(* IEC 61131-3 sources: daoli-st-library/DL_Process (part 51) *)

(* ---- FB_DL_ShiftHandoverCheck.st ---- *)
(*
  ==================================================================
  组件名 Component  : FB_DL_ShiftHandoverCheck
  分类   Category   : DL_Process
  复杂度 Complexity  : 中
  版本   Version    : 1.0.1
  功能   Purpose    : 班次交接检查。交接开始沿取运行快照（产量与报警计数），
                      交接窗 tHandover 内逐条确认未决事项，全部确认即置完成单拍
                      bHandoverDone；窗到期仍有未决项则升级故障码并转未完成态。
  来源   Source     : self-std（IEC 61131-3 标准时序 + 交接业务语义自研）
  溯源   Origin     : 班次交接检查为公开生产管理语义，道莅 clean-room 自研实现，
                      未复制任何厂商私有库源码。
  平台   Platform   : 纯 IEC 61131-3（TON / R_TRIG / 比较），三平台通用
  分工声明 Split     : 与 FB_DL_ShiftMonthReport（报表属主）与 FB_DL_ChangeoverSequence
                      （产品换型属主）双向互补——本件只做交接时点的检查与确认闭环，
                      不出报表、不做换型顺控、不改动生产计数本体。
  作者   Author     : 道莅代码库 · PLC 编程专家（R60）
  归属 Ownership     : E_DL_HandoverPhase 属主为本文件（全库唯一定义，R264）；
                      引用件只引用不重声明（D13 返修补行）。
  接口偏离声明       : nProdCnt / nAlarmCnt 为 UDINT 却沿用 n 前缀（D10 返修登记
                      例外，R200）：沿用派单既有引脚名不改，避免破坏调用方接口；
                      族内新件一律用 u 前缀。
  ------------------------------------------------------------------
  边界 Boundary     :
                      一 零长窗显式分支（R253）：tHandover ≤ 0 判组态非法故障码，
                         不进交接相（禁靠比较算子隐式分流）；
                      二 同拍竞态让位于合法事件（R275）：交汇段先消化本拍确认沿，
                         再消化窗口到期迁移——到期拍恰有确认沿时按确认处理，
                         不在同拍升级超窗码；
                      三 进入/退出条件逐条取反对偶（R259）：进入 = 开始沿 + 使能 +
                         窗合法 + 无锁存；退出 = 全确认（完成）/ 窗口到期（升级）/
                         失能（弃用）/ 复位沿（清锁存）四条并列；
                      四 快照「最近一次」类出口纳入复位清单（R243）：nSnapProd 与
                         nSnapAlarm 在复位沿一并清零；
                      五 单拍输出 bHandoverDone 统一出口段每拍先预置 FALSE、
                         分支只写 TRUE（R256）；
                      六 使能 bEnable = FALSE 时语义为「弃用本轮交接」（转空闲，
                         不锁存、不出单拍）——R191 声明行；
                      七 故障解除路径：eFault 相由复位沿迁回空闲并清锁存与快照
                         （bReset 为输入引脚，恒可达，R152 自证）。
  错误码   Codes    :
    16#0005_0620【信息级】交接窗内尚有未决事项（逐拍重算，不锁存）
    16#0005_0621【故障级】交接窗时长非法（≤0），组态非法，锁存至复位沿
    16#0005_0622【故障级】交接窗到期仍未全部确认，升级未完成故障，锁存至复位沿
  验收   Acceptance :
    算法已证（脚本）：未跑 ｜ 编译器已证（三平台）：未跑
    V1 3 项未决、窗内 3 个确认沿 → bHandoverDone 单拍、无故障
    V2 窗到期仅确认 2/3 → 码 0622、eFault、未完成
    V3 tHandover = T#0S → 首拍即码 0621，不进交接相
  修订记录 Revision  :
    2026-11-21  v1.0.0  R60 首版（批 3 · 序号 12）
    2026-11-21  v1.0.1  R61 返修：D7 增 _nPendingLock，仅 eIdle 迁入沿赋值，
                        判据与注释对齐（R259）；D10 n 前缀 UDINT 字段登记
                        例外；D13 补 E_DL_HandoverPhase 属主行
  ==================================================================
*)

TYPE E_DL_HandoverPhase :
(
    eIdle  := 0,  // 空闲：等交接开始沿 / idle, waiting for the start edge
    eWait  := 10, // 等待：交接窗内逐条确认 / waiting for the item confirmations inside the window
    eFault := 20  // 故障：窗非法或到期未完成，锁存待复位 / fault, an illegal window or an unfinished overrun, latched
);
END_TYPE

FUNCTION_BLOCK FB_DL_ShiftHandoverCheck
VAR_INPUT
    bEnable      : BOOL := TRUE;       // 使能，FALSE 时弃用本轮交接（边界六）/ the enable, false discards the round
    bStart       : BOOL := FALSE;      // 交接开始电平，上升沿取快照 / the start level, the rising edge takes the snapshot
    bConfirmItem : BOOL := FALSE;      // 未决事项确认电平，上升沿确认一条 / the item confirmation level, each rising edge confirms one item
    bReset       : BOOL := FALSE;      // 复位沿：清锁存与快照并回空闲 / the reset edge, clears the latch and the snapshot
    tHandover    : TIME := T#10M;      // 交接窗时长 [毫秒]，必须 > 0 / the handover window, must be positive
    nPendingItems : DINT := 3;         // 未决事项条数 [条]，合法域 0..64 / the pending item count, legal from zero to sixty four
    nProdCnt     : UDINT := 0;         // 当前班次产量计数 [件] / the production count of the shift
    nAlarmCnt    : UDINT := 0;         // 当前班次报警计数 [次] / the alarm count of the shift
END_VAR
VAR_OUTPUT
    bRunning       : BOOL := FALSE;               // 交接窗口进行中 [-] / the handover in progress flag
    bHandoverDone  : BOOL := FALSE;               // 交接完成单拍脉冲 [-] / the handover done one shot pulse
    nConfirmedCnt  : DINT := 0;                   // 已确认条数 [条] / the confirmed item count
    nSnapProd      : UDINT := 0;                  // 交接开始时刻的产量快照 [件] / the production snapshot at the start edge
    nSnapAlarm     : UDINT := 0;                  // 交接开始时刻的报警快照 [次] / the alarm snapshot at the start edge
    eState         : E_DL_HandoverPhase;          // 主状态机当前态 [状态] / the current state of the main machine
    bError         : BOOL := FALSE;               // 故障锁存位 [-] / the latched fault bit
    eErr           : UDINT := 16#0000_0000;       // 错误码，0 = 正常 / the error code, zero is ok
END_VAR
VAR
    _bInit      : BOOL := FALSE;                                 // 首拍初始化标志（R310）/ the first scan flag
    _eState     : E_DL_HandoverPhase := E_DL_HandoverPhase.eIdle; // 内部状态寄存器，段 4 唯一写点 / the internal state register, single writer
    _bDone      : BOOL := FALSE;                                 // 完成单拍内部位，段 1 预清段 6 映射 / the internal done bit, preset then mapped
    _nConfirmed : DINT := 0;                                     // 已确认条数副本 / the confirmed count copy
    _nPending   : DINT := 0;                                     // 未决条数钳位工作副本（逐拍重算，仅供迁入沿快照，D7 返修）/ the clamped pending work copy, recomputed every scan
    _nPendingLock : DINT := 0;                                   // 本轮未决条数锁定值（仅 eIdle 迁入沿赋值，D7 返修，R259）/ the locked pending count, assigned only on the idle entry edge
    _uSnapProd  : UDINT := 0;                                    // 产量快照副本 / the production snapshot copy
    _uSnapAlarm : UDINT := 0;                                    // 报警快照副本 / the alarm snapshot copy
    _bFault     : BOOL := FALSE;                                 // 故障锁存副本（仅复位沿清除）/ the fault latch copy
    _bCfgBad    : BOOL := FALSE;                                 // 组态非法标记（逐拍重算）[-] / the configuration fault flag
    _bIncomplete : BOOL := FALSE;                                // 未确认标记（逐拍重算）[-] / the unconfirmed flag
    rtStart     : R_TRIG;                                        // 开始沿实例，段 0 无条件刷新 / the start edge instance
    rtConfirm   : R_TRIG;                                        // 确认沿实例，段 0 无条件刷新 / the confirmation edge instance
    rtReset     : R_TRIG;                                        // 复位沿实例，段 0 无条件刷新 / the reset edge instance
    tonWindow   : TON;                                           // 交接窗定时器，段 0 无条件刷新 / the handover window timer
END_VAR
VAR CONSTANT
    DL_SHC_ITMAX : DINT := 64; // 未决事项上界 [条] / the pending item bound
END_VAR

// 段 0｜沿检测与交接窗定时器无条件周期刷新（禁入分支，R7；IN 串故障锁存门控，FB50-1）/ segment 0, the unconditional refresh with the latch gate
rtStart(CLK := bStart); // 开始沿 / the start edge
rtConfirm(CLK := bConfirmItem); // 确认沿 / the confirmation edge
rtReset(CLK := bReset); // 复位沿 / the reset edge
tonWindow(IN := (_eState = E_DL_HandoverPhase.eWait) AND (NOT _bFault), PT := tHandover); // 交接窗：仅等待相且无锁存时计时 / the window timing only in the waiting phase

// 段 1｜首拍初始化与单拍标志预清（仅单拍标志入清单，R32 FB32-1；R256）/ segment 1, the first scan init and the one shot preset
IF NOT _bInit THEN // 首拍一拍 / the first scan
    _bInit := TRUE; // 置首拍标志 / raise the first scan flag
    _nConfirmed := 0; // 已确认条数显式清零 / clear the confirmed count explicitly
    _nPending := 0; // 未决条数显式清零 / clear the pending count explicitly
    _nPendingLock := 0; // 未决锁定值显式清零（D7 返修）/ clear the locked pending count explicitly
    _uSnapProd := 0; // 产量快照显式清零 / clear the production snapshot explicitly
    _uSnapAlarm := 0; // 报警快照显式清零 / clear the alarm snapshot explicitly
    _bFault := FALSE; // 故障锁存显式清零 / clear the fault latch explicitly
    _eState := E_DL_HandoverPhase.eIdle; // 状态显式落空闲 / place the state to idle explicitly
END_IF
_bDone := FALSE; // 完成单拍预清零 / preset the done pulse false
_bCfgBad := FALSE; // 组态非法标记预清零 / preset the configuration flag false
_bIncomplete := FALSE; // 未确认标记预清零 / preset the unconfirmed flag false

// 段 2｜组态域闸（零长窗显式分支，边界一；未决条数越域钳位）/ segment 2, the configuration gate with the explicit zero length branch
IF tHandover <= T#0S THEN // 零长窗：非法组态 / a zero length window, an illegal configuration
    _bCfgBad := TRUE; // 置组态非法标记 / raise the configuration flag
    _bFault := TRUE; // 锁存故障（段 5 迁移相）/ latch the fault, the segment five migrates the phase
END_IF
IF nPendingItems < 0 THEN // 条目数为负（域下界硬限）/ a negative item count
    _nPending := 0; // 按零条处理（无未决即完成）/ treat as zero, an immediate completion
ELSIF nPendingItems > DL_SHC_ITMAX THEN // 条目数越上界 / above the bound
    _nPending := DL_SHC_ITMAX; // 钳到上界 / clamp to the bound
ELSE // 域内 / inside the domain
    _nPending := nPendingItems; // 原值接管 / take the value as is
END_IF

// 段 3｜本拍确认沿预消化（R275：合法事件先于窗口到期迁移消化，段序在段 4 之前）/ segment 3, the confirmation edge pre digest ahead of the window expiry
IF rtConfirm.Q AND (_eState = E_DL_HandoverPhase.eWait) AND (NOT _bFault) THEN // 等待相内的确认沿 / a confirmation edge inside the waiting phase
    IF _nConfirmed < _nPendingLock THEN // 尚有未确认条目（判据用锁定值，D7 返修）/ items remain unconfirmed against the locked count
        _nConfirmed := _nConfirmed + 1; // 确认一条 / confirm one item
    ELSE // 已全部确认（多按的确认沿忽略）/ everything is confirmed, extra presses ignored
        _nConfirmed := _nPendingLock; // 计数饱和于锁定条目数 / saturate the count at the locked item count
    END_IF
END_IF

// 段 4｜主状态机（ENUM + CASE，ELSE 拦非法态；进入/退出逐条取反对偶，边界三）/ segment 4, the main machine with the paired entry and exit conditions
CASE _eState OF
    E_DL_HandoverPhase.eIdle: // 空闲相：等开始沿（条件：开始沿 + 使能 + 窗合法 + 无锁存）/ the idle phase
        IF rtStart.Q AND bEnable AND (tHandover > T#0S) AND (NOT _bFault) THEN // 迁入判据带全量闸位复检（R274）/ the entry with the full gate recheck
            _nConfirmed := 0; // 新一轮确认计数归零 / reset the confirmed count
            _uSnapProd := nProdCnt; // 取产量快照（最近一次类出口）/ take the production snapshot
            _uSnapAlarm := nAlarmCnt; // 取报警快照 / take the alarm snapshot
            _nPendingLock := _nPending; // 未决条数锁定（仅此迁入沿赋值，窗内改参不影响本轮判据，D7 返修）/ lock the pending count on this entry edge only
            _eState := E_DL_HandoverPhase.eWait; // 迁入等待相 / enter the waiting phase
        END_IF
    E_DL_HandoverPhase.eWait: // 等待相：四条退出（全确认 / 到期 / 失能 / 锁存）/ the waiting phase with four exits
        IF _nConfirmed >= _nPendingLock THEN // 退出条件一：全部确认（判据用锁定值，D7 返修）/ the first exit, everything confirmed against the locked count
            _bDone := TRUE; // 置完成单拍 / raise the done pulse
            _eState := E_DL_HandoverPhase.eIdle; // 迁回空闲 / back to idle
        ELSIF tonWindow.Q THEN // 退出条件二：窗口到期仍未全部确认（边界二：本拍确认沿已在段 3 消化）/ the second exit, the window expired unconfirmed
            _bIncomplete := TRUE; // 置未确认标记 / raise the unconfirmed flag
            _bFault := TRUE; // 锁存超窗故障（0622）/ latch the overrun fault
        ELSIF (NOT bEnable) OR _bFault THEN // 退出条件三：失能弃用或已锁存（前置条件消失）/ the third exit with the prerequisite gone
            _eState := E_DL_HandoverPhase.eIdle; // 迁回空闲（不锁存、不出单拍）/ back to idle without a latch or a pulse
        END_IF
    E_DL_HandoverPhase.eFault: // 故障相：锁存保持，等复位沿（解除可达，边界七）/ the fault phase held until the reset edge
        IF rtReset.Q THEN // 复位沿（复位作用域：清锁存 + 清快照 + 清累计量 + 迁相位）/ the reset with the declared scope
            _bFault := FALSE; // 清故障锁存 / clear the fault latch
            _nConfirmed := 0; // 清确认计数 / clear the confirmed count
            _nPendingLock := 0; // 清未决锁定值（复位作用域含锁定值，D7 返修）/ clear the locked pending count within the reset scope
            _uSnapProd := 0; // 清产量快照（R243 最近一次类出口入复位清单）/ clear the production snapshot
            _uSnapAlarm := 0; // 清报警快照 / clear the alarm snapshot
            _eState := E_DL_HandoverPhase.eIdle; // 故障相迁出边回空闲 / the exit edge back to idle
        END_IF
    ELSE // 非法枚举值拦截 / the illegal enumeration guard
        _eState := E_DL_HandoverPhase.eIdle; // 落回空闲 / force back to idle
        _bFault := TRUE; // 置故障锁存 / latch the fault
END_CASE

// 段 5｜故障锁存迁移闸（置于解除段之后防同拍抢迁，R258）/ segment 5, the fault latch to phase gate placed after the release
IF _bFault AND (_eState <> E_DL_HandoverPhase.eFault) THEN // 已锁存但不在故障相 / latched but not in the fault phase
    _eState := E_DL_HandoverPhase.eFault; // 迁入故障相 / enter the fault phase
END_IF

// 段 6｜统一出口（内部副本单点映射，R180；故障码锁存回放，R187）/ segment 6, the unified outlet
_bIncomplete := (_eState = E_DL_HandoverPhase.eWait) AND (_nConfirmed < _nPendingLock); // 未确认提示逐拍重算（判据用锁定值，D7 返修）/ the unconfirmed hint recomputed every scan against the locked count
bRunning := (_eState = E_DL_HandoverPhase.eWait); // 进行中出口 / the in progress outlet
bHandoverDone := _bDone; // 完成单拍出口 / the done pulse outlet
nConfirmedCnt := _nConfirmed; // 确认条数出口 / the confirmed count outlet
nSnapProd := _uSnapProd; // 产量快照出口 / the production snapshot outlet
nSnapAlarm := _uSnapAlarm; // 报警快照出口 / the alarm snapshot outlet
eState := _eState; // 状态出口 / the state outlet
bError := _bFault; // 故障位出口（与锁存同源）/ the fault bit outlet from the same latch
IF _bFault THEN // 故障锁存回放优先 / the latched fault replays first
    IF _bCfgBad THEN // 组态成因（独立码值，R190）/ the configuration cause with its own code
        eErr := 16#0005_0621; // 故障级：交接窗时长非法 / fault grade, the window length is illegal
    ELSE // 超窗成因 / the overrun cause
        eErr := 16#0005_0622; // 故障级：到期仍未全部确认 / fault grade, still unconfirmed at the expiry
    END_IF
ELSIF _bIncomplete THEN // 未确认提示（信息级，逐拍重算）/ the informational unconfirmed hint
    eErr := 16#0005_0620; // 信息级：尚有未决事项 / informational, items still pending
    bError := FALSE; // 信息级不置 bError（仅故障级置位，R45 配对口径）/ the informational code never raises the fault bit
ELSE // 无事件 / no event
    eErr := 16#0000_0000; // 正常 / ok
END_IF
END_FUNCTION_BLOCK

(* ---- FB_DL_ShiftMonthReport.st ---- *)
(*
  ==================================================================
  组件名 Component  : FB_DL_ShiftMonthReport
  分类   Category   : DL_Process
  版本   Version    : 1.0.0
  功能   Purpose    : 班次 / 月度窗口产量报表闸。班次结束脉冲到达时结算本班产量
                      （好品 / 废品 / 良率）并累加进月度窗口，同时打开报表闸
                      （等上位确认或超时自动关闸），关闸拍出报表完成脉冲。
                      月变更沿清月度累计与班次计数，实现「班次窗 + 月度窗」双窗一致。
  溯源   Origin     : 班次 / 月度报表闸为通用产量统计语义；本件为 clean-room 实现，
                      仅借鉴来源分类与参数域组织（来源标签 roadmap-p2-shift），
                      道莅原创设计，未复制任何闭源代码行。
  平台   Platform   : 纯 IEC 61131-3（R_TRIG / TON / UDINT / REAL，无私有库）
  作者   Author     : 道莅代码库 · PLC 编程专家（R55）
  ------------------------------------------------------------------
  边界 Boundary     :
                      一 本件只做结算与报表闸控，不生成报表文件、不写数据库（属主边界）；
                      二 报表闸在「确认沿」或「闸超时」任一到达时关闭，两条路径均可达；
                      三 月度累计只在班次结算拍增长，禁按当下累计引脚每拍重算；
                      四 班次号越域与月变更属信息级事件，不置故障；
                      五 无全局变量、无外部变量声明、无物理地址寻址。
  输出契约 Output contract:
                      uShiftGood / uShiftScrap 为最近一次结算的班次量（锁存）；
                      uMonthGood / uMonthScrap 为当月累计（锁存，月变更清零）；
                      bReportDone 为单拍脉冲（内部位置位、统一出口映射后撤销）；
                      eCause 故障级成因与 bError 配对（R45），信息级永不置 bError。
  修订记录 Revision  :
    2026-11-20  v1.0.0  R55 首版（批 2 · 序号 8）
  ==================================================================
*)

TYPE E_DL_SmrState :
(
    eIdle   := 0,       // 空闲：等班次结束脉冲 / idle, waiting for the shift end pulse
    eGate   := 10,      // 报表闸开：等上位确认或闸超时 / report gate open, waiting for the acknowledgement or the gate timeout
    eFault  := 90       // 故障：组态非法锁存 / fault, illegal configuration latched
);
END_TYPE

TYPE E_DL_SmrCause :
(
    eNone       := 0,   // 无成因 / no cause
    eCfgIllegal := 1,   // 组态非法：月份、班次号或时间引脚越域（故障级，与 bError 配对）/ illegal config, month, shift index or time pin out of domain
    eShiftBad   := 2,   // 班次号越域已回钳（信息级）/ the shift index was clamped, informational
    eMonthRoll  := 3    // 月变更，月度累计已清零（信息级）/ month rolled over and the monthly accumulation was cleared, informational
);
END_TYPE

FUNCTION_BLOCK FB_DL_ShiftMonthReport
VAR_INPUT
    bEnable     : BOOL := TRUE;              // 使能，失能时关闸并冻结累计 [-] / enable, disabling closes the gate and freezes the accumulation
    bReset      : BOOL := FALSE;            // 复位上升沿清故障锁存与闸状态 [-] / reset rising edge clears the fault latch and the gate state
    nMonth      : INT := 1;                  // 当前月份 [月]，域 1..12 / current month [month], domain 1 to 12
    nShiftIdx   : INT := 1;                  // 当前班次号 [班]，域 1..3 / current shift index [shift], domain 1 to 3
    bShiftEnd   : BOOL := FALSE;             // 班次结束脉冲，上升沿结算 [-] / shift end pulse, settled on the rising edge
    uGoodCnt    : UDINT := 0;                // 本班好品累计 [只] / good pieces accumulated in the shift [pieces]
    uScrapCnt   : UDINT := 0;                // 本班废品累计 [只] / scrap pieces accumulated in the shift [pieces]
    bReportAck  : BOOL := FALSE;             // 上位确认报表，上升沿关闸 [-] / report acknowledgement, the rising edge closes the gate
    tGateTime   : TIME := T#30S;             // 报表闸超时 [毫秒]，域 大于零 / report gate timeout [millisecond], domain above zero
END_VAR
VAR_OUTPUT
    bReportGate : BOOL := FALSE;             // 报表闸开指示 [-] / report gate open indicator
    uShiftGood  : UDINT := 0;                // 最近结算班次好品数 [只] / good pieces of the last settled shift [pieces]
    uShiftScrap : UDINT := 0;                // 最近结算班次废品数 [只] / scrap pieces of the last settled shift [pieces]
    fShiftYield : REAL := 0.0;               // 最近结算班次良率 [百分比] / yield of the last settled shift [percent]
    uMonthGood  : UDINT := 0;                // 当月好品累计 [只] / monthly good pieces [pieces]
    uMonthScrap : UDINT := 0;                // 当月废品累计 [只] / monthly scrap pieces [pieces]
    fMonthYield : REAL := 0.0;               // 当月良率 [百分比] / monthly yield [percent]
    nMonthShifts: INT := 0;                  // 当月已结算班次数 [班] / settled shifts within the month [shift]
    bReportDone : BOOL := FALSE;             // 报表完成单拍脉冲 [-] / report done single-shot pulse
    eState      : E_DL_SmrState := E_DL_SmrState.eIdle; // 相位出口 [枚举] / phase outlet [enum]
    eCause      : E_DL_SmrCause := E_DL_SmrCause.eNone; // 成因出口 [枚举] / cause outlet [enum]
    bError      : BOOL := FALSE;             // 故障锁存标志 [-] / fault latch flag
END_VAR
VAR
    rtShift     : R_TRIG;                    // 班次结束沿检测，段 0 无条件刷新 / shift end edge detector, refreshed unconditionally in segment zero
    rtAck       : R_TRIG;                    // 报表确认沿检测，段 0 无条件刷新 / acknowledgement edge detector, refreshed unconditionally in segment zero
    rtReset     : R_TRIG;                    // 复位沿检测，段 0 无条件刷新 / reset edge detector, refreshed unconditionally in segment zero
    tonGate     : TON;                       // 报表闸超时，段 0 无条件刷新 / report gate timeout, refreshed unconditionally in segment zero
    _eState     : E_DL_SmrState := E_DL_SmrState.eIdle;  // 内部相位，CASE 唯一写入目标 / internal phase, the only CASE write target
    _eCause     : E_DL_SmrCause := E_DL_SmrCause.eNone;  // 信息级成因，每拍重算 / informational cause, recomputed every scan
    _eFaultCause: E_DL_SmrCause := E_DL_SmrCause.eNone;  // 故障级成因，锁存至复位沿 / fault cause, latched until the reset edge
    _bFault     : BOOL := FALSE;             // 故障锁存位 [-] / fault latch bit
    _bInit      : BOOL := FALSE;             // 首扫初始化完成标志（R310）/ first scan initialisation flag
    _bDoneInt   : BOOL := FALSE;             // 报表完成脉冲内部位，统一出口映射 / internal done bit, mapped at the unified outlet
    _bShiftBad  : BOOL := FALSE;             // 班次号被回钳 [-] / the shift index was clamped
    _bCfgBad    : BOOL := FALSE;             // 组态非法判定 [-] / illegal configuration verdict
    _bYieldOk   : BOOL := FALSE;             // 良率除子可用 [-] / the yield divisor is usable
    _nMonthPrev : INT := -1;                 // 上一拍月份快照，初值 -1 使首拍必清 / previous month snapshot, minus one forces a clear on the first scan
    _nShiftUse  : INT := 1;                  // 钳定后的班次号 [班] / clamped shift index [shift]
    _uGoodLoc   : UDINT := 0;                // 本拍好品暂存 [只] / good pieces held in a local [pieces]
    _uScrapLoc  : UDINT := 0;                // 本拍废品暂存 [只] / scrap pieces held in a local [pieces]
    _uMonthG    : UDINT := 0;                // 当月好品累加器 [只] / monthly good accumulator [pieces]
    _uMonthS    : UDINT := 0;                // 当月废品累加器 [只] / monthly scrap accumulator [pieces]
    _uShiftG    : UDINT := 0;                // 班次好品保持块 [只] / shift good holder [pieces]
    _uShiftS    : UDINT := 0;                // 班次废品保持块 [只] / shift scrap holder [pieces]
    _uTotLoc    : UDINT := 0;                // 良率分母（好品加废品）[只] / yield denominator, good plus scrap [pieces]
    _uMonthTot  : UDINT := 0;                // 月度良率分母（好品加废品）[只] / monthly yield denominator [pieces]
    _fYield     : REAL := 0.0;               // 良率工作值 [百分比] / yield working value [percent]
END_VAR
VAR CONSTANT
    DL_SMR_SHIFT_MIN : INT := 1;             // 班次号下限 [班] / shift index floor [shift]
    DL_SMR_SHIFT_MAX : INT := 3;             // 班次号上限 [班] / shift index ceiling [shift]
    DL_SMR_CNT_MAX   : UDINT := 2147483647;  // 计数加和上限，防 UDINT 相加溢出后窄化 [只] / summation ceiling against overflow before narrowing [pieces]
    DL_SMR_YIELD_MAX : REAL := 100.0;        // 良率上限 [百分比] / yield ceiling [percent]
    DL_SMR_DAY_SHIFT_MAX : INT := 3;         // 单日班次计数的自然上限 [班] / natural ceiling of the daily shift count [shift]
END_VAR

// 段 0｜定时器与沿检测无条件周期刷新（禁入分支），IN 只串状态闸 / segment 0, unconditional refresh of timers and edges with state gates on IN only
rtShift(CLK := bShiftEnd); // 班次结束沿无条件刷新 / unconditional refresh of the shift end edge
rtAck(CLK := bReportAck); // 确认沿无条件刷新 / unconditional refresh of the acknowledgement edge
rtReset(CLK := bReset); // 复位沿无条件刷新 / unconditional refresh of the reset edge
tonGate(IN := (_eState = E_DL_SmrState.eGate) AND (NOT _bFault), PT := tGateTime); // 报表闸超时，IN 串相位闸与故障闸 / report gate timeout with the phase gate and the fault gate on IN

// 段 1｜首扫初始化（R310）/ segment 1, first scan initialisation
IF NOT _bInit THEN // 首扫一拍 / the very first scan
    _bInit := TRUE; // 置首扫完成标志 / raise the first scan flag
    _eState := E_DL_SmrState.eIdle; // 相位从空闲起步 / the phase starts from idle
    _eCause := E_DL_SmrCause.eNone; // 信息级成因清零 / clear the informational cause
    _eFaultCause := E_DL_SmrCause.eNone; // 故障级成因清零 / clear the fault cause
    _bFault := FALSE; // 故障锁存清零 / clear the fault latch
    _nMonthPrev := -1; // 月份快照置非法值 / put the month snapshot at an illegal value
    _uMonthG := 0; // 月度好品清零 / clear monthly good pieces
    _uMonthS := 0; // 月度废品清零 / clear monthly scrap pieces
    nMonthShifts := 0; // 月度班次计数清零 / clear the monthly shift count
END_IF

// 段 2｜复位沿作用域：清锁存 / 迁相位 / 清闸内部位（累计不清，避免产量丢失）/ segment 2, reset edge scope
IF rtReset.Q THEN // 复位沿 / reset edge
    _bFault := FALSE; // 作用域一：清故障锁存 / scope one, clear the fault latch
    _eFaultCause := E_DL_SmrCause.eNone; // 作用域一：清故障级成因 / scope one, clear the fault cause
    _eState := E_DL_SmrState.eIdle; // 作用域二：迁回空闲相 / scope two, migrate back to idle
    _bDoneInt := FALSE; // 作用域二：清完成脉冲内部位 / scope two, clear the internal done bit
    _eCause := E_DL_SmrCause.eNone; // 作用域一：清信息级成因 / scope one, clear the informational cause
END_IF

// 段 3｜组态域闸（R151 全覆盖）/ segment 3, configuration domain gate over every pin
_bCfgBad := FALSE; // 组态非法预置假 / preset the illegal configuration verdict to false
IF (nMonth < 1) OR (nMonth > 12) THEN // 月份越域 / month out of domain
    _bCfgBad := TRUE; // 判非法 / mark illegal
END_IF
IF (nShiftIdx < DL_SMR_SHIFT_MIN) OR (nShiftIdx > DL_SMR_SHIFT_MAX) THEN // 班次号越域 / shift index out of domain
    _bCfgBad := TRUE; // 判非法 / mark illegal
END_IF
IF tGateTime <= T#0S THEN // 闸超时非正 / gate timeout not positive
    _bCfgBad := TRUE; // 判非法 / mark illegal
END_IF
IF _bCfgBad AND (NOT _bFault) THEN // 组态非法且未锁存 / illegal configuration and not yet latched
    _bFault := TRUE; // 置故障锁存 / raise the fault latch
    _eFaultCause := E_DL_SmrCause.eCfgIllegal; // 故障级成因 (R45 配对 bError) / fault grade cause paired with bError
    _eState := E_DL_SmrState.eFault; // 迁故障相 / migrate to the fault phase
END_IF
_nShiftUse := nShiftIdx; // 班次号直通 / shift index passes through
_bShiftBad := FALSE; // 回钳标志预置假 / preset the clamp flag to false
IF _nShiftUse < DL_SMR_SHIFT_MIN THEN // 下越界 / below the lower bound
    _nShiftUse := DL_SMR_SHIFT_MIN; // 回钳到 1 / clamp to one
    _bShiftBad := TRUE; // 置回钳标志 / raise the clamp flag
ELSIF _nShiftUse > DL_SMR_SHIFT_MAX THEN // 上越界 / above the upper bound
    _nShiftUse := DL_SMR_SHIFT_MAX; // 回钳到 3 / clamp to three
    _bShiftBad := TRUE; // 置回钳标志 / raise the clamp flag
END_IF

// 段 4｜月变更：清月度累计与班次计数（信息级事件，不置故障）/ segment 4, month rollover clears the monthly accumulation, an informational event
_eCause := E_DL_SmrCause.eNone; // 信息级成因每拍重算 / the informational cause is recomputed every scan
IF (nMonth <> _nMonthPrev) THEN // 月份变化（首拍必命中）/ month changed, always true on the first scan
    _nMonthPrev := nMonth; // 月份快照推进 / advance the month snapshot
    _uMonthG := 0; // 月度好品清零 / clear monthly good pieces
    _uMonthS := 0; // 月度废品清零 / clear monthly scrap pieces
    nMonthShifts := 0; // 月度班次计数清零 / clear the monthly shift count
    _uShiftG := 0; // 班次保持块清零 / clear the shift holder
    _uShiftS := 0; // 班次保持块清零 / clear the shift holder
    _eCause := E_DL_SmrCause.eMonthRoll; // 信息级成因：月变更已清零 / informational cause, the rollover cleared the accumulation
END_IF
IF _bShiftBad THEN // 班次号被回钳 / the shift index was clamped
    _eCause := E_DL_SmrCause.eShiftBad; // 信息级成因覆盖（同拍仅报更具体者）/ the informational cause overrides for the more specific event
END_IF

// 段 5｜相位机：ENUM + CASE，含 ELSE 非法相位兜底（R128）/ segment 5, phase machine with an ELSE fallback for illegal phases
CASE _eState OF
E_DL_SmrState.eIdle: // 空闲相：等班次结束脉冲 / idle phase, waiting for the shift end pulse
    IF rtShift.Q AND (NOT _bFault) THEN // 班次结束沿且无故障 / shift end edge without a fault
        _uGoodLoc := uGoodCnt; // 好品暂存 / hold the good pieces
        _uScrapLoc := uScrapCnt; // 废品暂存 / hold the scrap pieces
        _uTotLoc := _uGoodLoc + _uScrapLoc; // 良率分母 / yield denominator
        IF (_uTotLoc < _uGoodLoc) OR (_uTotLoc < _uScrapLoc) THEN // 相加回绕 / the sum wrapped around
            _uTotLoc := DL_SMR_CNT_MAX; // 饱和到上限，防窄化负值（R316 口径）/ saturated at the ceiling against a negative narrowing
        END_IF
        _bYieldOk := _uTotLoc > 0; // 分母可用性 / denominator usability
        IF _bYieldOk THEN // 分母可用 / the denominator is usable
            _fYield := UDINT_TO_REAL(_uGoodLoc) / UDINT_TO_REAL(_uTotLoc) * 100.0; // 良率，除子已证大于零 / yield, divisor proven positive
            IF _fYield > DL_SMR_YIELD_MAX THEN // 良率越上限 / yield above the ceiling
                _fYield := DL_SMR_YIELD_MAX; // 上钳 / clamp upward
            END_IF
        ELSE
            _fYield := 0.0; // 无产量时良率记零 / zero yield when nothing was produced
        END_IF
        _uShiftG := _uGoodLoc; // 班次好品保持 / hold the shift good pieces
        _uShiftS := _uScrapLoc; // 班次废品保持 / hold the shift scrap pieces
        IF (_uMonthG + _uGoodLoc) < _uMonthG THEN // 累加回绕 / the accumulation wrapped around
            _uMonthG := DL_SMR_CNT_MAX; // 饱和到上限 / saturated at the ceiling
        ELSE
            _uMonthG := _uMonthG + _uGoodLoc; // 月度好品累加 / accumulate monthly good pieces
        END_IF
        IF (_uMonthS + _uScrapLoc) < _uMonthS THEN // 累加回绕 / the accumulation wrapped around
            _uMonthS := DL_SMR_CNT_MAX; // 饱和到上限 / saturated at the ceiling
        ELSE
            _uMonthS := _uMonthS + _uScrapLoc; // 月度废品累加 / accumulate monthly scrap pieces
        END_IF
        IF nMonthShifts < DL_SMR_DAY_SHIFT_MAX THEN // 班次计数未越自然上限 / the shift count is below its natural ceiling
            nMonthShifts := nMonthShifts + 1; // 班次计数递增 / increment the shift count
        END_IF
        _eState := E_DL_SmrState.eGate; // 迁报表闸相 / migrate to the report gate phase
    END_IF

E_DL_SmrState.eGate: // 报表闸相：确认沿或闸超时关闸 / report gate phase, closed by the acknowledgement edge or the gate timeout
    IF rtAck.Q OR tonGate.Q THEN // 确认或超时 / acknowledged or timed out
        _bDoneInt := TRUE; // 报表完成脉冲内部位置位（统一出口映射，R187）/ raise the internal done bit, mapped at the unified outlet
        _eState := E_DL_SmrState.eIdle; // 迁回空闲相 / migrate back to idle
    END_IF

E_DL_SmrState.eFault: // 故障相：锁存回放，等复位沿 / fault phase, the latch is replayed until the reset edge
    _bDoneInt := FALSE; // 故障拍不出完成脉冲 / no done pulse while faulted

ELSE // 非法相位兜底（R128）/ illegal phase fallback
    _bFault := TRUE; // 置故障锁存 / raise the fault latch
    _eFaultCause := E_DL_SmrCause.eCfgIllegal; // 故障级成因记组态非法 / record the illegal configuration cause
    _eState := E_DL_SmrState.eFault; // 迁故障相 / migrate to the fault phase
END_CASE

// 段 6｜失能语义：关闸并冻结累计（R191 显式声明）/ segment 6, disabled semantics, close the gate and freeze the accumulation
IF NOT bEnable THEN // 失能 / disabled
    _eState := E_DL_SmrState.eIdle; // 迁回空闲相 / migrate back to idle
    _bDoneInt := FALSE; // 撤完成脉冲内部位 / withdraw the internal done bit
END_IF

// 段 7｜统一出口 / segment 7, unified outlet
bReportGate := (_eState = E_DL_SmrState.eGate); // 闸开指示（挂状态量）/ gate open indicator as a state quantity
uShiftGood := _uShiftG; // 班次好品出口 / shift good outlet
uShiftScrap := _uShiftS; // 班次废品出口 / shift scrap outlet
fShiftYield := _fYield; // 班次良率出口 / shift yield outlet
uMonthGood := _uMonthG; // 月度好品出口 / monthly good outlet
uMonthScrap := _uMonthS; // 月度废品出口 / monthly scrap outlet
_uMonthTot := _uMonthG + _uMonthS; // 月度分母先落局部量，避免重复计算 / the monthly denominator lands in a local first
IF _uMonthTot < _uMonthG THEN // 相加回绕 / the sum wrapped around
    _uMonthTot := DL_SMR_CNT_MAX; // 饱和到上限 / saturated at the ceiling
END_IF
IF _uMonthTot > 0 THEN // 月度分母可用 / the monthly denominator is usable
    fMonthYield := UDINT_TO_REAL(_uMonthG) / UDINT_TO_REAL(_uMonthTot) * 100.0; // 月度良率，除子已证大于零 / monthly yield, divisor proven positive
    IF fMonthYield > DL_SMR_YIELD_MAX THEN // 良率越上限 / yield above the ceiling
        fMonthYield := DL_SMR_YIELD_MAX; // 上钳 / clamp upward
    END_IF
ELSE
    fMonthYield := 0.0; // 无产量时良率记零 / zero yield when nothing was produced
END_IF
eState := _eState; // 相位出口单点映射 / single-point phase outlet mapping
bReportDone := _bDoneInt; // 完成脉冲映射本拍值 / map the done pulse for this scan
_bDoneInt := FALSE; // 映射后立即撤销，保证单拍宽度（R187 两段式）/ revoke right after mapping to keep a single-scan width
IF _bFault THEN // 故障锁存优先 / the fault latch takes priority
    eCause := _eFaultCause; // 故障级成因锁存回放 / the fault cause is replayed from the latch
ELSE
    eCause := _eCause; // 信息级成因直映 / the informational cause is mapped directly
END_IF
bError := _bFault; // 故障标志与锁存位同源 / the fault flag shares the latch source
END_FUNCTION_BLOCK

(* ---- FB_DL_ShrinkTunnelCtrl.st ---- *)
(*
  FB_DL_ShrinkTunnelCtrl  —  热收缩炉温区-网速联动三段工艺窗 / Shrink tunnel zone-temperature to belt-speed linkage in three process windows
  分类 Category : DL_Process
  版本 Version  : 1.0.0
  来源 Source   : t1-2-oscat — 工艺联动族零检索深化
  溯源 Origin   : clean-room 实现，未复制任何源码行
  功能 Function : 1) 三段配方顺控：ePre（预缩）→ eMain（主缩）→ eSettle（定型）→ eDone，
                  段推进 TON（tonAdvPre/tonAdvMain/tonAdvSet）与总超时 TON（tonPhaseTo）
                  成对分实例（R233 纪律）；
                  2) 温区-网速联动：温区均温（来源 = 上游 FB_DL_HeatCoolZone 各区温度镜像，
                  经 aZoneTemp 引脚注入，本件不实例化 HeatCoolZone——每区需四重接口注入，
                  组合方式见边界①）落当前段窗 [fXxxLo, fXxxHi] → 网速设定 = fVelMax；
                  越窗 → 降速至 fVelMin（保窗优先），越窗沿/回窗沿置信息级；
                  3) 段推进沿 048F；越窗降速激活沿 0490；回窗恢复沿 0491；
                  4) 段超时或非法相位兜底 → 0369 锁存；温度非有限 → 0368 锁存。
  边界 Boundary : ① 温度源组合方式：上游每温区一个 FB_DL_HeatCoolZone 实例，其加热/冷却
                  执行后的区温（或经 I_DL_AnalogSensor 读数）由调用方逐区镜像入 aZoneTemp；
                  本件只消费温度数值做工艺窗判定，不承载温区 PID（分工：HeatCoolZone 管区
                  内恒温，本件管跨区工艺窗与网速联动）；
                  ② 组态闸：uZoneCnt < 1 或 > 8、fVelMin <= 0 或 >= fVelMax、任一窗上下限
                  颠倒 → 0367 锁存；
                  ③ 网速下限 > 0 组态闸（防零速死锁）；配方推进与超时 TON 分实例；
                  ④ 无 GVL 依赖：纯引脚输入输出，无外部变量引用，无物理 IO 地址。
  依赖 Depends  : 与 FB_DL_HeatCoolZone 温度镜像组合（不实例化）；Standard.library（TON / R_TRIG）
  码表 Error codes（Process 段 0005，窗口 0367~0369 / 048F~0491）:
    16#0005_0367 故障级：组态非法（站数/网速域/工艺窗颠倒），锁存至 bReset
    16#0005_0368 故障级：温区温度非有限（NaN 自反判），锁存至 bReset
    16#0005_0369 故障级：段超时或相位落 ELSE 兜底，锁存至 bReset
    16#0005_048F 信息级：段推进沿（Pre→Main→Settle）
    16#0005_0490 信息级：越窗降速激活沿
    16#0005_0491 信息级：回窗恢复沿（降速解除）
  修订历史 Revision :
    2026-11-19  v1.0.0  R41 首版（批次 4 · 序号 3）
*)

TYPE E_DL_ShrinkPhase :
(
    eIdle   := 0,    // 空闲：等启动沿 / Idle, waiting start edge
    ePre    := 10,   // 预缩段 / Pre-shrink phase
    eMain   := 20,   // 主缩段 / Main-shrink phase
    eSettle := 30,   // 定型段 / Settle phase
    eDone   := 40,   // 完成 / Done
    eFault  := 90    // 故障 / Fault
);
END_TYPE

FUNCTION_BLOCK FB_DL_ShrinkTunnelCtrl
VAR_INPUT
    aZoneTemp    : ARRAY[1..8] OF LREAL;  // 各温区实际温度 [°C]（HeatCoolZone 镜像）/ Zone temperatures mirrored
    uZoneCnt     : UINT := 1;         // 温区数 [区]，域 1..8 / Zone count
    fVelMin      : LREAL := 5.0;      // 网速下限（降速保窗档）[m/min]，域 > 0 / Belt speed lower bound
    fVelMax      : LREAL := 30.0;     // 网速正常档 [m/min]，域 > fVelMin / Belt speed normal bound
    fPreLo       : LREAL := 120.0;    // 预缩窗下限 [°C] / Pre-shrink window low
    fPreHi       : LREAL := 160.0;    // 预缩窗上限 [°C] / Pre-shrink window high
    fMainLo      : LREAL := 180.0;    // 主缩窗下限 [°C] / Main-shrink window low
    fMainHi      : LREAL := 220.0;    // 主缩窗上限 [°C] / Main-shrink window high
    fSetLo       : LREAL := 90.0;     // 定型窗下限 [°C] / Settle window low
    fSetHi       : LREAL := 130.0;    // 定型窗上限 [°C] / Settle window high
    tPreDur      : TIME := T#30S;     // 预缩段时长 [ms]，域 > 0 / Pre-phase duration
    tMainDur     : TIME := T#60S;     // 主缩段时长 [ms]，域 > 0 / Main-phase duration
    tSetDur      : TIME := T#45S;     // 定型段时长 [ms]，域 > 0 / Settle-phase duration
    tTotalTo     : TIME := T#300S;    // 配方总超时 [ms]，域 > 0 / Total recipe timeout
    bStart       : BOOL := FALSE;     // 启动沿 [-] / Start edge
    bReset       : BOOL := FALSE;     // 复位，上升沿清故障锁存 / Reset edge clears fault latch
END_VAR
VAR_OUTPUT
    ePhase       : E_DL_ShrinkPhase;  // 段出口，段尾单点映射 / Phase outlet
    fVelSet      : LREAL;             // 网速设定出口 [m/min] / Belt speed setpoint outlet
    bTempOk      : BOOL;              // 温度落当前段窗标志 [-] / Temperature in-window flag
    bError       : BOOL;              // 故障锁存标志 / Fault latch flag
    nErrId       : UDINT;             // 事件码，0 = 无事件 / Event code
END_VAR
VAR
    tonAdvPre    : TON;               // 预缩段推进 TON，无条件刷新 / Pre-phase advance timer
    tonAdvMain   : TON;               // 主缩段推进 TON，无条件刷新 / Main-phase advance timer
    tonAdvSet    : TON;               // 定型段推进 TON，无条件刷新 / Settle-phase advance timer
    tonPhaseTo   : TON;               // 配方总超时 TON（专用超时命名），无条件刷新 / Total timeout timer
    rtStart      : R_TRIG;            // 启动沿实例，无条件刷新 / Start edge instance
    rtReset      : R_TRIG;            // 复位沿实例，无条件刷新 / Reset edge instance
    _eState      : E_DL_ShrinkPhase := E_DL_ShrinkPhase.eIdle;  // 内部相位（CASE 唯一写入目标）/ Internal phase
    _fZoneAvg    : LREAL;             // 温区均温 [°C] / Zone average temperature
    _nCap        : INT;               // 生效温区数 [区] / Effective zone count
    _bInWin      : BOOL;              // 温度落窗当拍量 [-] / In-window current-scan flag
    _bSlowPrev   : BOOL;              // 上拍降速镜像（回窗沿判据）/ Previous slow mirror
    _bFault      : BOOL;              // 故障锁存位（锁存量）/ Latched fault bit
    _uFault      : UDINT;             // 故障码锁存（锁存量）/ Latched fault code
    _uInfo       : UDINT;             // 信息码，每拍重算 / Transient info code
    i            : INT;               // 均温循环游标 [索引] / Average loop cursor
    _nGuard      : INT;               // 均温守卫计数 [次] / Average guard counter
END_VAR

(* —— 段 0：定时器与沿实例无条件周期刷新（禁置于 IF/CASE 内） —— *)
rtStart(CLK := bStart);                                   // 启动沿（每拍必调）
rtReset(CLK := bReset);                                   // 复位沿（每拍必调）
tonAdvPre(IN := (_eState = E_DL_ShrinkPhase.ePre), PT := tPreDur);      // 预缩推进（单相独占）
tonAdvMain(IN := (_eState = E_DL_ShrinkPhase.eMain), PT := tMainDur);   // 主缩推进（单相独占）
tonAdvSet(IN := (_eState = E_DL_ShrinkPhase.eSettle), PT := tSetDur);   // 定型推进（单相独占）
tonPhaseTo(IN := (_eState = E_DL_ShrinkPhase.ePre)
           OR (_eState = E_DL_ShrinkPhase.eMain)
           OR (_eState = E_DL_ShrinkPhase.eSettle), PT := tTotalTo);    // 总超时（配方相集合）

(* —— 段 1：单拍量预清零（锁存量 _bFault/_uFault 不入清单，禁同拍抹除） —— *)
_uInfo := 16#0000_0000;             // 信息码每拍重算
nErrId := 16#0000_0000;             // 事件码缺省无事件

(* —— 段 2：复位沿 + 组态域闸（当拍量判据；网速下限 > 0 组态闸） —— *)
IF rtReset.Q THEN                   // rtReset.Q = 当拍量
    _bFault := FALSE;               // 清故障锁存位
    _uFault := 16#0000_0000;        // 清故障锁存码
    _eState := E_DL_ShrinkPhase.eIdle;  // 相位回空闲
END_IF
_nCap := UINT_TO_INT(uZoneCnt);     // 温区数快照
IF (_nCap < 1) OR (_nCap > 8) OR (fVelMin <= 0.0) OR (fVelMin >= fVelMax)
   OR (fPreLo >= fPreHi) OR (fMainLo >= fMainHi) OR (fSetLo >= fSetHi)
   OR (TIME_TO_DINT(tTotalTo) <= 0) THEN
    _uFault := 16#0005_0367;        // 故障级：组态非法
    _bFault := TRUE;
END_IF

(* —— 段 3：温区均温计算（LREAL 口径；守卫循环；防除零由 uZoneCnt 组态闸承载） —— *)
_fZoneAvg := 0.0;                   // 均温累加器清零
_nGuard := 0;                       // 守卫清零
IF (NOT _bFault) AND (_nCap >= 1) AND (_nCap <= 8) THEN
    FOR i := 1 TO _nCap DO
        _nGuard := _nGuard + 1;     // 守卫递增
        IF _nGuard > 8 THEN
            EXIT;                   // 守卫兜底退出（理论不可达）
        END_IF
        IF (aZoneTemp[i] <> aZoneTemp[i]) OR ((aZoneTemp[i] - aZoneTemp[i]) <> (aZoneTemp[i] - aZoneTemp[i])) THEN
            _uFault := 16#0005_0368;    // 故障级：温区温度非有限
            _bFault := TRUE;
        END_IF
        _fZoneAvg := _fZoneAvg + aZoneTemp[i];  // 累加
    END_FOR
    IF NOT _bFault THEN
        _fZoneAvg := _fZoneAvg / INT_TO_LREAL(_nCap);   // 均温（分母 >= 1 已过闸，防除零）
    END_IF
END_IF

(* —— 段 4：工艺窗判定与网速联动（当拍量判据） —— *)
CASE _eState OF
E_DL_ShrinkPhase.ePre:
    _bInWin := (_fZoneAvg >= fPreLo) AND (_fZoneAvg <= fPreHi);     // 预缩窗判定
E_DL_ShrinkPhase.eMain:
    _bInWin := (_fZoneAvg >= fMainLo) AND (_fZoneAvg <= fMainHi);   // 主缩窗判定
E_DL_ShrinkPhase.eSettle:
    _bInWin := (_fZoneAvg >= fSetLo) AND (_fZoneAvg <= fSetHi);     // 定型窗判定
ELSE
    _bInWin := FALSE;               // 非工艺相无窗判定
END_CASE
bTempOk := _bInWin AND (NOT _bFault);   // 落窗出口
IF (NOT _bFault) AND bStart THEN
    IF _bInWin THEN
        fVelSet := fVelMax;         // 落窗：正常档网速
        IF _bSlowPrev THEN
            _uInfo := 16#0005_0491; // 信息级：回窗恢复沿
        END_IF
    ELSE
        fVelSet := fVelMin;         // 越窗：降速保窗
        IF NOT _bSlowPrev THEN
            _uInfo := 16#0005_0490; // 信息级：越窗降速激活沿
        END_IF
    END_IF
ELSE
    fVelSet := 0.0;                 // 非运行相网速归零（安全侧）
END_IF

(* —— 段 5：配方相位机（CASE 全覆盖 + ELSE 兜底） —— *)
CASE _eState OF

E_DL_ShrinkPhase.eIdle:
    IF rtStart.Q AND (NOT _bFault) THEN
        _eState := E_DL_ShrinkPhase.ePre;   // 进预缩段
    END_IF

E_DL_ShrinkPhase.ePre:
    IF _bFault THEN
        _eState := E_DL_ShrinkPhase.eFault; // 故障相
    ELSIF tonPhaseTo.Q THEN
        _uFault := 16#0005_0369;            // 故障级：配方总超时
        _bFault := TRUE;
        _eState := E_DL_ShrinkPhase.eFault;
    ELSIF tonAdvPre.Q THEN
        _uInfo := 16#0005_048F;             // 信息级：段推进沿
        _eState := E_DL_ShrinkPhase.eMain;  // 进主缩段
    END_IF

E_DL_ShrinkPhase.eMain:
    IF _bFault THEN
        _eState := E_DL_ShrinkPhase.eFault; // 故障相
    ELSIF tonPhaseTo.Q THEN
        _uFault := 16#0005_0369;            // 故障级：配方总超时
        _bFault := TRUE;
        _eState := E_DL_ShrinkPhase.eFault;
    ELSIF tonAdvMain.Q THEN
        _uInfo := 16#0005_048F;             // 信息级：段推进沿
        _eState := E_DL_ShrinkPhase.eSettle;    // 进定型段
    END_IF

E_DL_ShrinkPhase.eSettle:
    IF _bFault THEN
        _eState := E_DL_ShrinkPhase.eFault; // 故障相
    ELSIF tonPhaseTo.Q THEN
        _uFault := 16#0005_0369;            // 故障级：配方总超时
        _bFault := TRUE;
        _eState := E_DL_ShrinkPhase.eFault;
    ELSIF tonAdvSet.Q THEN
        _uInfo := 16#0005_048F;             // 信息级：段推进沿
        _eState := E_DL_ShrinkPhase.eDone;  // 进完成相
    END_IF

E_DL_ShrinkPhase.eDone:
    IF NOT bStart THEN
        _eState := E_DL_ShrinkPhase.eIdle;  // 指令撤销回空闲
    END_IF

E_DL_ShrinkPhase.eFault:
    ;                                   // 故障相：等复位沿（段 2 承载迁出）

ELSE
    _uFault := 16#0005_0369;            // 故障级：非法相位兜底（归并超时码，头注释码表声明）
    _bFault := TRUE;
    _eState := E_DL_ShrinkPhase.eFault; // 强制回故障相

END_CASE

(* —— 段 6：出口单点映射（名实同源；锁存码回放，禁同拍抹除） —— *)
IF _bFault THEN
    nErrId := _uFault;              // 故障锁存码回放
    fVelSet := 0.0;                 // 故障期网速归零（安全侧）
    bTempOk := FALSE;               // 故障期落窗出口 FALSE（安全侧）
ELSE
    nErrId := _uInfo;               // 信息码
END_IF
bError := _bFault;                  // 故障标志与锁存位同源
ePhase := _eState;                  // 状态出口单点映射
_bSlowPrev := (NOT _bInWin) AND (NOT _bFault);   // 降速镜像快照

END_FUNCTION_BLOCK

(* ---- FB_DL_SiloLevelInterlock.st ---- *)
// =====================================================================
// FB_DL_SiloLevelInterlock.st
// 料仓高低料位-输送联锁（防溢仓/空跑双联锁 + 卡料窗）
// Silo level interlock with conveyor, overflow/empty trips and jam window
// 所属子库: DL_Process    版本: v1.0.0    兼容: CODESYS V3.5+ / TwinCAT 3 / 汇川 InoProShop
// 码位: 16#0005_046C ~ 16#0005_0470 (本件独占 5 槽, 勿复用)
// 溯源: 道莅 clean-room 防御性实现
//       来源组标签: process-control, silo, interlock, conveyor
// 修改记录: R30 初版 (ROUND_PLAN_R30 序 7)
// 安全声明: 料位开关以假 = 未到达该料位为正常态（失电安全侧: 开关失电判为
//           未到达）; 输送允许输出安全侧为假; 各锁存位解除式均可达
// =====================================================================
FUNCTION_BLOCK FB_DL_SiloLevelInterlock
VAR_INPUT
    bHighLevel : BOOL := FALSE;     // 高料位开关, 真 = 到达高料位 / High level switch, TRUE = reached
    bLowLevel  : BOOL := FALSE;     // 低料位开关, 真 = 到达低料位 / Low level switch, TRUE = reached
    bConvRun   : BOOL := FALSE;     // 输送运行反馈 / Conveyor run feedback
    bRunDemand : BOOL := FALSE;     // 输送运行需求注入（上位流程给出, 供卡料判据使用）/ Run demand injected
    tJamWin    : TIME := T#5S;      // 卡料确认窗 T#100MS~T#60S / Jam confirm window [s]
    bReset     : BOOL := FALSE;     // 联锁复位命令 / Interlock reset command
END_VAR
VAR_OUTPUT
    bConvPermit   : BOOL := FALSE;  // 输送允许, 安全侧为假; 高料位联锁只停进料不停输送 / Conveyor permit, safe FALSE
    bOverflowTrip : BOOL := FALSE;  // 溢仓联锁锁存 / Overflow trip latch
    bEmptyTrip    : BOOL := FALSE;  // 空跑联锁锁存 / Empty-run trip latch
    bJamDet       : BOOL := FALSE;  // 卡料检测锁存 / Jam detection latch
    eErr          : UDINT := 16#0005_046C;  // 错误码 / Error code
END_VAR
VAR
    rtrReset  : R_TRIG;             // 复位上升沿检测, 每拍无条件刷新 / Reset edge, refreshed every cycle
    tonJam    : TON;                // 卡料确认定时器, 每拍无条件刷新 / Jam confirm timer, refreshed every cycle
    bConflict : BOOL := FALSE;      // 料位组态矛盾锁存 / Level configuration conflict latch
END_VAR

// ---------------------------------------------------------------------
// 代码位表（本件独占, 勿复用）:
//   16#0005_046C 信息 联锁正常（输送允许且无锁存事件）
//   16#0005_046D 故障 料位组态矛盾（高低料位同时有效）,
//                解除式 = 双开关恢复互斥 且 bReset 上升沿
//   16#0005_046E 故障 溢仓联锁（高料位: 停进料, 输送允许保持完成当前批次）,
//                解除式 = 高料位消失 且 bReset 上升沿
//   16#0005_046F 故障 空跑联锁（低料位: 停输送防空跑）,
//                解除式 = 低料位消失 且 bReset 上升沿
//   16#0005_0470 故障 卡料（运行需求持续而输送无反馈超窗）,
//                解除式 = 输送反馈恢复 且 bReset 上升沿
// ---------------------------------------------------------------------

// ---- 复位沿实例无条件刷新 / Unconditional reset edge refresh ----
rtrReset(CLK := bReset);

// ---- 组态矛盾与联锁锁存置位（锁存置位, 解除见各解除式）/ Conflict and trip latches ----
IF bHighLevel AND bLowLevel THEN
    bConflict := TRUE;              // 高低料位同时有效 = 组态矛盾 / Both levels active = conflict
END_IF
IF bHighLevel THEN
    bOverflowTrip := TRUE;          // 高料位置溢仓联锁 / High level sets overflow trip
END_IF
IF bLowLevel THEN
    bEmptyTrip := TRUE;             // 低料位置空跑联锁 / Low level sets empty trip
END_IF

// ---- 卡料确认定时器无条件周期刷新（有运行需求而无运行反馈才计时）/ Jam timer unconditional refresh ----
tonJam(IN := bRunDemand AND (NOT bConvRun) AND (NOT bJamDet)
        AND (NOT bConflict) AND (NOT bEmptyTrip),
       PT := tJamWin);
IF tonJam.Q THEN
    bJamDet := TRUE;                // 窗内持续无反馈判卡料 / No feedback through window = jam
END_IF

// ---- 锁存解除式（全部可达, R28 自证）/ Latch release paths, all reachable ----
IF rtrReset.Q AND (NOT (bHighLevel AND bLowLevel)) THEN
    bConflict := FALSE;             // 矛盾解除: 双开关恢复互斥 / Conflict release
END_IF
IF rtrReset.Q AND (NOT bHighLevel) THEN
    bOverflowTrip := FALSE;         // 溢仓解除: 高料位消失 / Overflow release
END_IF
IF rtrReset.Q AND (NOT bLowLevel) THEN
    bEmptyTrip := FALSE;            // 空跑解除: 低料位消失 / Empty release
END_IF
IF rtrReset.Q AND bConvRun THEN
    bJamDet := FALSE;               // 卡料解除: 运行反馈恢复 / Jam release
END_IF

// ---- 输送允许: 矛盾/空跑/卡料任一锁存即禁止; 溢仓联锁不停输送（完成当前批次）
//      Conveyor permit: blocked by conflict/empty/jam; overflow keeps conveyor ----
bConvPermit := (NOT bConflict) AND (NOT bEmptyTrip) AND (NOT bJamDet);

// ---- 错误码仲裁（联锁动作与告警码分离输出）/ Error arbitration ----
IF bConflict THEN
    eErr := 16#0005_046D;           // 组态矛盾 / Configuration conflict
ELSIF bOverflowTrip THEN
    eErr := 16#0005_046E;           // 溢仓联锁 / Overflow trip
ELSIF bEmptyTrip THEN
    eErr := 16#0005_046F;           // 空跑联锁 / Empty trip
ELSIF bJamDet THEN
    eErr := 16#0005_0470;           // 卡料 / Jam
ELSE
    eErr := 16#0005_046C;           // 联锁正常 / Interlock normal
END_IF

END_FUNCTION_BLOCK

(* ---- FB_DL_SinterFurnaceRampCtrl.st ---- *)
(*
  Component : FB_DL_SinterFurnaceRampCtrl
  Category  : DL_Process
  Type      : FB
  Complexity: C2
  VERSION   : v1.0.0
  功能      : 烧结炉升温曲线跟踪：ENUM 七态（Idle/Purge/Ramp/Soak/Cool/Done/Fault），斜率限幅给定值输出，露点超限联锁，吹扫/保温/冷却分段计时。
  开源溯源  : 道莅原创 clean-room 自研（无外部代码引用）｜License: MIT
  边界条件  : ① 升温斜率、目标温度、露点上限、各段时长为判据基，须 > 1e-9 或非 0，否则拒启动并锁故障；
              ② 给定值斜率限幅按采样周期积分推进（每个采样节拍最多走 斜率×dt/60），禁阶跃；
              ③ 露点超上限在吹扫/升温/保温三相均联锁，故障锁存唯一解除路径 = bReset 上升沿。
*)

TYPE E_DL_SintPhase :
(
    eIdle  := 0,    (* 空闲：等启动沿 / Idle waiting start edge *)
    ePurge := 10,   (* 吹扫：露点置换 / Atmosphere purge *)
    eRamp  := 20,   (* 升温：斜率限幅跟踪 / Ramp with slope limit *)
    eSoak  := 30,   (* 保温：目标温度保持 / Soak at target *)
    eCool  := 40,   (* 冷却：斜率限幅下降 / Controlled cooling *)
    eDone  := 50,   (* 完成：曲线结束 / Curve finished *)
    eFault := 90    (* 故障：锁存待复位 / Fault latched *)
);
END_TYPE

FUNCTION_BLOCK FB_DL_SinterFurnaceRampCtrl
VAR_INPUT
    bEnable    : BOOL;   (* 使能电平 [-] Enable level *)
    bReset     : BOOL;   (* 复位上升沿，清故障锁存 [-] Reset edge *)
    bStart     : BOOL;   (* 启动上升沿 [-] Start edge *)
    fActC      : REAL;   (* 炉膛实测温度 [°C] Measured furnace temperature *)
    fTargetC   : REAL;   (* 目标保温温度 [°C] Target soaking temperature *)
    fCoolToC   : REAL;   (* 冷却终点温度 [°C] Cooling end temperature *)
    fRampCmin  : REAL;   (* 允许升温/降温斜率 [°C/min] Allowed ramp rate *)
    fDewPointC : REAL;   (* 炉内实测露点 [°C] Measured dew point *)
    fDewMaxC   : REAL;   (* 露点允许上限 [°C] Dew point upper limit *)
    tPurge     : TIME;   (* 吹扫驻留 [ms] Purge dwell *)
    tSoak      : TIME;   (* 保温驻留 [ms] Soak dwell *)
    tCool      : TIME;   (* 冷却超时保护 [ms] Cooling timeout *)
    tSample    : TIME;   (* 斜率积分采样周期 [ms] Ramp integration period *)
END_VAR
VAR_OUTPUT
    fSetOutC : REAL;              (* 温度给定值输出 [°C] Temperature setpoint output *)
    bHeatOn  : BOOL;              (* 加热使能输出 [-] Heater enable output *)
    ePhase   : E_DL_SintPhase;    (* 相位出口，段尾单点映射 [-] Phase outlet *)
    bError   : BOOL;              (* 故障锁存标志 [-] Fault latch flag *)
    uErrId   : UDINT;             (* 事件码，0 = 无事件 [-] Event code *)
END_VAR
VAR
    rtReset  : R_TRIG;   (* 复位沿实例，每拍无条件刷新 / Reset edge *)
    rtStart  : R_TRIG;   (* 启动沿实例，每拍无条件刷新 / Start edge *)
    tonPurge : TON;      (* 吹扫驻留计时（独立实例） / Purge timer *)
    tonSoak  : TON;      (* 保温驻留计时（独立实例） / Soak timer *)
    tonCool  : TON;      (* 冷却计时（独立实例） / Cooling timer *)
    tonSample: TON;      (* 采样节拍（自复位错峰） / Sampling tick self-reset *)
    _ePhase  : E_DL_SintPhase := E_DL_SintPhase.eIdle;  (* 内部相位 / Internal phase *)
    _bFault  : BOOL;     (* 故障锁存位（锁存量） / Latched fault bit *)
    _uFault  : UDINT;    (* 故障码锁存（锁存量） / Latched fault code *)
    _bCfgBad : BOOL;     (* 组态非法当拍量 [-] Config illegal flag *)
    _bNonFin : BOOL;     (* 输入非有限当拍量 [-] Non-finite input flag *)
    fDt      : REAL;     (* 采样周期秒值 [s] Sampling period in seconds *)
    fStepK   : REAL;     (* 单拍允许最大温度变化量 [K] Max temperature step per tick *)
END_VAR
VAR CONSTANT
    DL_EPS      : REAL := 1.0E-9;   (* 除零判定容差 [无量纲] Divide-by-zero tolerance *)
    DL_MS_PER_S : REAL := 1000.0;   (* 毫秒转秒换算系数 [ms/s] Milliseconds per second *)
    DL_S_PER_MIN: REAL := 60.0;     (* 分钟转秒换算系数 [s/min] Seconds per minute *)
    DL_ZERO     : REAL := 0.0;      (* 零常量 [无量纲] Zero constant *)
END_VAR

(* —— 段 0｜沿与定时器每拍无条件刷新（禁置于 IF/CASE 内，使能挂 IN 引脚） —— *)
rtReset(CLK := bReset);
rtStart(CLK := bStart);
tonPurge (IN := (_ePhase = E_DL_SintPhase.ePurge) AND (NOT _bFault), PT := tPurge);
tonSoak  (IN := (_ePhase = E_DL_SintPhase.eSoak)  AND (NOT _bFault), PT := tSoak);
tonCool  (IN := (_ePhase = E_DL_SintPhase.eCool)  AND (NOT _bFault), PT := tCool);
tonSample(IN := NOT tonSample.Q, PT := tSample);

(* —— 段 1｜每拍量预清零（锁存量 _bFault/_uFault/fSetOutC 不入清单） —— *)
uErrId := 16#0000_0000;
_bCfgBad := FALSE;
_bNonFin := FALSE;
bHeatOn := FALSE;

(* —— 段 2｜复位沿：故障一次性清干净，给定值跟随实测，相位回空闲 —— *)
IF rtReset.Q THEN
    _bFault := FALSE;
    _uFault := 16#0000_0000;
    fSetOutC := fActC;
    _ePhase := E_DL_SintPhase.eIdle;
END_IF

(* —— 段 3｜非有限拦截与组态闸（覆盖斜率/目标/露点/各段时长） —— *)
IF (fActC <> fActC) OR ((fActC - fActC) <> 0.0)
   OR (fTargetC <> fTargetC) OR ((fTargetC - fTargetC) <> 0.0)
   OR (fDewPointC <> fDewPointC) OR ((fDewPointC - fDewPointC) <> 0.0)
   OR (fRampCmin <> fRampCmin) OR ((fRampCmin - fRampCmin) <> 0.0)
   OR (fCoolToC <> fCoolToC) OR ((fCoolToC - fCoolToC) <> 0.0) THEN
    _bNonFin := TRUE;
END_IF
IF (fRampCmin <= DL_EPS) OR (fDewMaxC = DL_ZERO) OR (tPurge = T#0S)
   OR (tSoak = T#0S) OR (tCool = T#0S) OR (tSample = T#0S) THEN
    _bCfgBad := TRUE;
END_IF

(* —— 段 4｜斜率限幅单拍步长：每个采样节拍最多走 斜率 × dt / 60 —— *)
fDt := TIME_TO_REAL(tSample) / DL_MS_PER_S;
fStepK := fRampCmin * fDt / DL_S_PER_MIN;

(* —— 段 5｜主状态机：七态全覆盖 + ELSE 兜底 —— *)
CASE _ePhase OF
E_DL_SintPhase.eIdle:
    fSetOutC := fActC;                       (* 空闲：给定跟随实测，无加热 *)
    IF rtStart.Q AND bEnable AND (NOT _bFault) AND (NOT _bCfgBad) AND (NOT _bNonFin) THEN
        _ePhase := E_DL_SintPhase.ePurge;
    ELSIF rtStart.Q AND (_bFault OR _bCfgBad OR _bNonFin) THEN
        _bFault := TRUE;                     (* 带病启动拒绝 / Reject start with bad config *)
        _uFault := 16#0027_0001;
        _ePhase := E_DL_SintPhase.eFault;
    END_IF

E_DL_SintPhase.ePurge:
    fSetOutC := fActC;                       (* 吹扫相不升温 *)
    IF (_bNonFin) OR (fDewPointC > fDewMaxC) THEN
        _bFault := TRUE; _uFault := 16#0027_0002;   (* 故障级：露点超限/输入非有限 *)
        _ePhase := E_DL_SintPhase.eFault;
    ELSIF tonPurge.Q THEN
        _ePhase := E_DL_SintPhase.eRamp;            (* 迁出条件 1：吹扫驻留完成 *)
    ELSIF NOT bEnable THEN
        _ePhase := E_DL_SintPhase.eIdle;            (* 迁出条件 2：使能撤销回安全态 *)
    END_IF

E_DL_SintPhase.eRamp:
    bHeatOn := TRUE;
    (* 给定值按单拍步长向目标推进，禁阶跃（斜率限幅） *)
    IF tonSample.Q THEN
        IF (fTargetC - fSetOutC) > fStepK THEN
            fSetOutC := fSetOutC + fStepK;
        ELSIF (fSetOutC - fTargetC) > fStepK THEN
            fSetOutC := fSetOutC - fStepK;
        ELSE
            fSetOutC := fTargetC;
        END_IF
    END_IF
    IF (_bNonFin) OR (fDewPointC > fDewMaxC) THEN
        _bFault := TRUE; _uFault := 16#0027_0002;   (* 故障级：露点超限/输入非有限 *)
        _ePhase := E_DL_SintPhase.eFault;
    ELSIF (fTargetC - fSetOutC) <= (fStepK + DL_EPS) THEN
        _ePhase := E_DL_SintPhase.eSoak;            (* 迁出条件 1：到达保温温度 *)
    ELSIF NOT bEnable THEN
        _ePhase := E_DL_SintPhase.eIdle;            (* 迁出条件 2：使能撤销 *)
    END_IF

E_DL_SintPhase.eSoak:
    bHeatOn := TRUE;
    fSetOutC := fTargetC;                    (* 保温相给定恒为目标温度 *)
    IF (_bNonFin) OR (fDewPointC > fDewMaxC) THEN
        _bFault := TRUE; _uFault := 16#0027_0002;   (* 故障级：露点超限/输入非有限 *)
        _ePhase := E_DL_SintPhase.eFault;
    ELSIF tonSoak.Q THEN
        _ePhase := E_DL_SintPhase.eCool;            (* 迁出条件 1：保温驻留完成 *)
    ELSIF NOT bEnable THEN
        _ePhase := E_DL_SintPhase.eIdle;            (* 迁出条件 2：使能撤销 *)
    END_IF

E_DL_SintPhase.eCool:
    (* 冷却相给定按单拍步长下降，加热输出撤销 *)
    IF tonSample.Q THEN
        IF (fSetOutC - fCoolToC) > fStepK THEN
            fSetOutC := fSetOutC - fStepK;
        ELSE
            fSetOutC := fCoolToC;
        END_IF
    END_IF
    IF tonCool.Q THEN
        _bFault := TRUE; _uFault := 16#0027_0003;   (* 故障级：冷却超时 *)
        _ePhase := E_DL_SintPhase.eFault;
    ELSIF fSetOutC <= (fCoolToC + DL_EPS) THEN
        _ePhase := E_DL_SintPhase.eDone;            (* 迁出条件 1：达冷却终点 *)
    ELSIF NOT bEnable THEN
        _ePhase := E_DL_SintPhase.eIdle;            (* 迁出条件 2：使能撤销 *)
    END_IF

E_DL_SintPhase.eDone:
    bHeatOn := FALSE;
    IF NOT bStart THEN
        _ePhase := E_DL_SintPhase.eIdle;            (* 启动撤销：回空闲 *)
    END_IF

E_DL_SintPhase.eFault:
    bHeatOn := FALSE;                        (* 故障相：加热输出安全侧撤销 *)

ELSE
    _bFault := TRUE;                         (* 兜底：非法相位锁存 *)
    _uFault := 16#0027_0009;
    _ePhase := E_DL_SintPhase.eFault;
END_CASE

(* —— 段 6｜相位与故障码出口单点映射 —— *)
ePhase := _ePhase;
bError := _bFault;
IF _bFault AND (_uFault <> 16#0000_0000) THEN
    uErrId := _uFault;                       (* 故障码锁存回放 / Latched fault replay *)
END_IF
END_FUNCTION_BLOCK

(* ---- FB_DL_SlurryDensityTrim.st ---- *)
(*==============================================================================
 * 组件名称 (Component)  : FB_DL_SlurryDensityTrim
 * 所属子库 (Sublibrary) : DL_Process
 * 当前版本 (Version)    : 1.0.0
 * 兼容性 (Platform)     : CODESYS 3.5+ / TwinCAT 3 / 汇川 InoProShop / 施耐德 Machine Expert
 *                         仅依赖 Standard.library（TON / R_TRIG / ABS），零厂商私有库
 * 功能描述 (Function)   : 浆料面密度双源交叉校核与分档告警。负载式与 β 射线
 *                         两路面密度源求均值出出面密度，双源偏差超容差持续
 *                         tMisDly 即 bMismatch 告警（防单拍毛刺）；均值对工艺
 *                         窗 [fBandLo, fBandHi] 分档 eLow/eIn/eHigh。与
 *                         ToleranceWindow（单源判窗）分工：本件是多源一致性
 *                         新判据 + 分档告警。
 * 来源标签 (Origin)     : ROADMAP §16.1 R11 池（L695），自研 clean-room
 * 边界语义 (Boundary)   : ① 双源任一非有限拍：冻结（均值/判档保持上拍，不告
 *                         警不消警）；
 *                         ② 一致性容差/窗界域闸（fBandLo < fBandHi）→ 组态故障；
 *                         ③ 告警去抖 TON 电平计时（非自复位周期窗）。
 * 输出语义 (Fallback)   : 【R191】bEnable = FALSE → 均值/分档保持末值 + 告警
 *                         收敛 FALSE（失能必须收敛告警）；eFault 相 → 冻结
 *                         + bError = TRUE。
 * 码位     (Codes)      : 按 R297 范式零 16# 码位硬编码；错误出口 BOOL+ENUM(eCause)。
 * 红线自检 (Redline)    : 7 项红线已自检：R1 零全局 ✓｜R2 零物理地址 ✓｜R3 纯 IEC ✓
 *                         R4 除零无涉/NaN 冻结/组态闸 ✓｜R5 双语同行注释 ✓
 *                         R6 CASE 带 ELSE 兜底迁 eFault ✓｜R7 TON/R_TRIG 段 0 无条件刷新 ✓
 * 验收向量 (Acceptance) : V1 双源 98.0/98.2（容差 0.5）→ 均值 98.1，
 *                         窗 [95,105] → eGrade=eIn，bMismatch=FALSE；
 *                         V2 双源 98.0/100.9（偏差 2.9 > 0.5）持续 tMisDly
 *                         → bMismatch=TRUE；
 *                         V3 均值 94.0 < 95 → eGrade=eLow，bAlarmLo=TRUE。
 * 修订历史 (Revision)   : 2026-11-20  v1.0.0  R51 首版（批 1 · 序号 4）
 *==============================================================================*)
TYPE E_DL_SdtGrade :
(
    eLow  := 0,                              (* 低于工艺窗 / Below window *)
    eIn   := 1,                              (* 窗内合格 / In window *)
    eHigh := 2                               (* 高于工艺窗 / Above window *)
);
END_TYPE

TYPE E_DL_SdtState :
(
    eIdle  := 0,                             (* 待使能 / Idle *)
    eRun   := 10,                            (* 双源校核运行 / Cross-check run *)
    eFault := 90                             (* 故障锁存相 / Fault latched phase *)
);
END_TYPE

TYPE E_DL_SdtCause :
(
    eNone       := 0,                        (* 无故障成因 / No cause *)
    eCfgIllegal := 1,                        (* 组态非法：窗界倒置/容差越域 / Illegal config *)
    ePhaseBad   := 2                         (* 非法相位兜底 / Illegal phase fallback *)
);
END_TYPE

FUNCTION_BLOCK FB_DL_SlurryDensityTrim
VAR_INPUT
    fDenLoad   : LREAL := 0.0;               (* 负载式面密度源 1 [g/m²] / Loadcell areal density *)
    fDenBeta   : LREAL := 0.0;               (* β 射线面密度源 2 [g/m²] / Beta-gauge areal density *)
    fBandLo    : LREAL := 95.0;              (* 工艺窗下限，域 < fBandHi [g/m²] / Window lower bound *)
    fBandHi    : LREAL := 105.0;             (* 工艺窗上限，域 > fBandLo [g/m²] / Window upper bound *)
    fTolPair   : LREAL := 0.5;               (* 双源一致性容差，域 > 0 [g/m²] / Cross-source tolerance *)
    tMisDly    : TIME := T#2S;               (* 失配告警去抖时长，域 > T#0S [ms] / Mismatch debounce *)
    bEnable    : BOOL := TRUE;               (* 使能 [-] / Enable *)
    bReset     : BOOL := FALSE;              (* 复位命令，上升沿清全部 [-] / Reset command *)
END_VAR
VAR_OUTPUT
    fDenAvg    : LREAL;                      (* 双源均值出面密度 [g/m²] / Averaged density *)
    eGrade     : E_DL_SdtGrade;              (* 分档出口 / Grade outlet *)
    bMismatch  : BOOL;                       (* 双源失配告警（去抖后电平）[-] / Mismatch alarm *)
    bAlarmLo   : BOOL;                       (* 低档告警电平 [-] / Low alarm *)
    bAlarmHi   : BOOL;                       (* 高档告警电平 [-] / High alarm *)
    eState     : E_DL_SdtState;              (* 状态出口 / State outlet *)
    eCause     : E_DL_SdtCause;              (* 故障成因出口 / Fault cause outlet *)
    bError     : BOOL;                       (* 故障锁存标志 [-] / Fault latch flag *)
END_VAR
VAR
    _eState  : E_DL_SdtState := E_DL_SdtState.eIdle;      (* 内部相位（CASE 唯一写入目标） / Internal phase *)
    _eCause  : E_DL_SdtCause := E_DL_SdtCause.eNone;      (* 故障成因锁存量 / Latched cause *)
    rtReset  : R_TRIG;                       (* 复位沿实例，段 0 无条件调用 / Reset edge instance *)
    tonMis   : TON;                          (* 失配去抖计时，段 0 无条件调用 / Mismatch debounce *)
    _fAvg    : LREAL;                        (* 均值派生量 [g/m²] / Average derived *)
    _bSrcBad : BOOL;                         (* 双源非有限当拍量 [-] / Non-finite source *)
    _bMisRaw : BOOL;                         (* 失配原始判据电平 [-] / Raw mismatch level *)
    _bFault  : BOOL;                         (* 故障锁存位 / Latched fault bit *)
    _bCfgBad : BOOL;                         (* 组态非法当拍量 / Illegal config this scan *)
END_VAR
VAR CONSTANT
    DL_SDT_EPS : LREAL := 1.0E-9;            (* 容差判零容差 [g/m²] / Tolerance epsilon *)
END_VAR

(* —— 段 0：当拍判据派生 + 实例无条件刷新（R228A） —— *)
_bCfgBad := (fTolPair <= DL_SDT_EPS) OR (fBandLo >= fBandHi) OR (tMisDly <= T#0S);   (* 组态闸（R151 全引脚 + 窗界序） / Config gate *)
rtReset(CLK := bReset);                      (* 复位沿每拍必调 / Reset edge every scan *)
_bSrcBad := (fDenLoad <> fDenLoad) OR ((fDenLoad - fDenLoad) <> (fDenLoad - fDenLoad))
            OR (fDenBeta <> fDenBeta) OR ((fDenBeta - fDenBeta) <> (fDenBeta - fDenBeta));   (* 双源 NaN 自反 + Inf 差判 / Non-finite source gates *)
tonMis(IN := (_eState = E_DL_SdtState.eRun) AND (NOT _bSrcBad) AND _bMisRaw, PT := tMisDly);   (* 失配去抖（电平计时非周期窗） / Mismatch debounce *)

(* —— 段 1：单拍量预清零（R107） —— *)
_fAvg := 0.0;                                (* 均值预清（每拍全路径派生，R285） / Average preset *)
_bMisRaw := FALSE;                           (* 失配原始判据预清 / Raw mismatch preset *)
bAlarmLo := FALSE;                           (* 低档告警预清（全路径赋值） / Low alarm preset *)
bAlarmHi := FALSE;                           (* 高档告警预清 / High alarm preset *)
eGrade := E_DL_SdtGrade.eIn;                 (* 分档缺省窗内（判定分支覆盖） / Grade preset *)

(* —— 段 2：复位沿处理（作用域：清故障 + 清均值出口 + 清分档 + 迁 eIdle，R283 逐项声明） —— *)
IF rtReset.Q THEN
    _bFault := FALSE;                        (* 清故障锁存 / Clear fault *)
    _eCause := E_DL_SdtCause.eNone;          (* 清成因 / Clear cause *)
    fDenAvg := 0.0;                          (* 清均值出口 / Clear average outlet *)
    eGrade := E_DL_SdtGrade.eIn;             (* 分档复位窗内 / Grade reset *)
    _eState := E_DL_SdtState.eIdle;          (* 迁待机相 / Back to idle *)
END_IF

(* —— 段 3：组态闸故障锁存（R45 配对；锁存至复位沿，R189） —— *)
IF _bCfgBad AND NOT _bFault THEN
    _bFault := TRUE;                         (* 锁存故障位 / Latch fault *)
    _eCause := E_DL_SdtCause.eCfgIllegal;    (* 成因：组态非法 / Cause: illegal config *)
    _eState := E_DL_SdtState.eFault;         (* 同步迁故障相 / Migrate to fault *)
END_IF

(* —— 段 4：CASE 主状态机（ELSE 兜底迁 eFault，红线 6） —— *)
CASE _eState OF
    E_DL_SdtState.eIdle:                     (* 待机相 / Idle *)
        IF bEnable AND NOT _bFault AND NOT _bSrcBad THEN
            _eState := E_DL_SdtState.eRun;   (* 进入运行 / Enter run *)
        END_IF
    E_DL_SdtState.eRun:                      (* 运行相：均值 + 失配 + 分档 / Run *)
        IF NOT bEnable THEN
            bMismatch := FALSE;              (* 失能告警收敛（R191 声明） / Alarm converge on disable *)
            _eState := E_DL_SdtState.eIdle;  (* 回待机 / Back to idle *)
        ELSIF NOT _bSrcBad THEN
            _fAvg := 0.5 * (fDenLoad + fDenBeta);   (* 双源均值（除子常量 2，无除零） / Average *)
            fDenAvg := _fAvg;                (* 均值出口刷新 / Average outlet *)
            _bMisRaw := ABS(fDenLoad - fDenBeta) > fTolPair;   (* 失配原始判据（容差闸） / Raw mismatch *)
            bMismatch := tonMis.Q;           (* 去抖后告警出口 / Debounced alarm *)
            IF _fAvg < fBandLo THEN
                eGrade := E_DL_SdtGrade.eLow;   (* 低档 / Low *)
            ELSIF _fAvg > fBandHi THEN
                eGrade := E_DL_SdtGrade.eHigh;  (* 高档 / High *)
            ELSE
                eGrade := E_DL_SdtGrade.eIn;    (* 窗内（IF 链带 ELSE 兜底，R285） / In window *)
            END_IF
            bAlarmLo := (eGrade = E_DL_SdtGrade.eLow) AND (NOT bMismatch);   (* 低档告警（失配时双源不可信不判档告警，R146 方向拆分） / Low alarm *)
            bAlarmHi := (eGrade = E_DL_SdtGrade.eHigh) AND (NOT bMismatch);  (* 高档告警 / High alarm *)
        END_IF                               (* 源坏值拍：冻结保持（边界①），告警不消不增 / Bad source: freeze *)
    E_DL_SdtState.eFault:                    (* 故障相：冻结保持，仅复位沿出 / Fault *)
        bMismatch := FALSE;                  (* 故障相告警收敛（安全侧） / Alarm converge in fault *)
    ELSE                                     (* 非法相位兜底迁安全态 / Illegal phase fallback *)
        _eState := E_DL_SdtState.eFault;     (* 迁故障相 / To fault *)
        _bFault := TRUE;                     (* 同步锁存 / Latch *)
        _eCause := E_DL_SdtCause.ePhaseBad;  (* 成因：非法相位 / Cause: illegal phase *)
END_CASE

(* —— 段 5：出口映射（bError/eState 同源，R191） —— *)
bError := _bFault;                           (* 故障标志镜像 / Fault flag mirror *)
eState := _eState;                           (* 状态出口 / State outlet *)
eCause := _eCause;                           (* 成因出口 / Cause outlet *)
END_FUNCTION_BLOCK

(* ---- FB_DL_SlurrySieveClogWatch.st ---- *)
(*
  ==================================================================
  组件名 Component  : FB_DL_SlurrySieveClogWatch
  分类   Category   : DL_Process
  复杂度 Complexity  : cx4
  版本   Version    : 1.0.0
  功能   Purpose    : 浆料筛网堵塞监视。堵塞指数 = (dP / q²) 对学习基准的比值；
                      趋势斜率取时间序环窗 8 点（R194：时间序遍历，禁头游标序）
                      最小二乘斜率；劣化分 warn / alarm 双级独立成因（R190）；
                      流量低于下限判 eFlowLoss；基准仅在清洁态持续窗口内更新。
  来源   Source     : t2-6-rockwell-aoi（判据组织次源）
  溯源   Origin     : IEC 61131-3 标准语义的道莅防御性实现；压差 / 流量堵塞判据为
                      公开过滤工艺语义，clean-room 自研实现，未复制任何闭源代码行。
  平台   Platform   : 纯 IEC 61131-3（TON / R_TRIG / ARRAY / LREAL，无私有库）
  作者   Author     : 道莅代码库 · PLC 编程专家（R56）
  ------------------------------------------------------------------
  边界 Boundary     :
                      一 本件只做堵塞判级与基准学习，不反冲洗、不调流量（属主边界）；
                      二 环窗遍历一律按时间序（自最旧样本起，R194）；最小二乘分母
                         8·Σx² - (Σx)² = 8·140 - 784 = 336，x = 0..7 结构性非零；
                      三 判据方向性（R146）：warn 与 alarm 为同向递进双级，成因独立；
                      四 学习判据：严重度 < fCleanRatio 持续 tLearnWin 才更新基准
                         （rtLearn 边沿单次更新，防每拍重写）；
                      五 成因锁存解除路径 = 迟滞反向自愈 或 bReset 上升沿（R188）；
                      六 无全局变量、无外部变量声明、无物理地址寻址。
  输出契约 Output contract:
                      fClogIdx 为堵塞指数（相对基准，1.0 = 基准水平）；fTrendSlope 为
                      8 点最小二乘斜率（每拍）；eFault 为锁存回放；
                      ePhaseBad 为非法相位兜底专用成员（R128）。
  修订记录 Revision  :
    2026-11-20  v1.0.0  R56 首版（批 3 · 序号 15）
  ==================================================================
*)

TYPE E_DL_SscPhase :
(
    eIdle  := 0,  // 未使能：监视停摆 / disabled, the watch is idle
    eRun   := 10, // 运行：逐拍判级 / running, graded every scan
    eFault := 90  // 故障：成因锁存 / fault, the cause is latched
);
END_TYPE

TYPE E_DL_SscFault :
(
    eNone      := 0, // 无成因 / no cause
    eClogWarn  := 1, // 堵塞预警级（故障级，与 bError 配对）/ the clog warning grade, fault grade paired with bError
    eClogAlarm := 2, // 堵塞报警级（故障级，与 bError 配对）/ the clog alarm grade, fault grade paired with bError
    eFlowLoss  := 3, // 流量低于下限（故障级，与 bError 配对）/ the flow is below the floor, fault grade paired with bError
    eSensorBad := 4, // 压差或流量非有限（故障级，与 bError 配对）/ the pressure or the flow is non finite, fault grade paired with bError
    ePhaseBad  := 5  // 非法相位兜底（故障级，与 bError 配对）/ illegal phase fallback, fault grade paired with bError
);
END_TYPE

FUNCTION_BLOCK FB_DL_SlurrySieveClogWatch
VAR_INPUT
    bEnable     : BOOL := TRUE;   // 使能，失能时监视停摆 [-] / enable, the watch stops when disabled
    bReset      : BOOL := FALSE;  // 复位上升沿清全部锁存与环窗 [-] / reset rising edge clears every latch and the ring
    fDp         : LREAL := 10.0;  // 筛前筛后压差 [千帕] / the sieve differential pressure [kilopascal]
    fQ          : LREAL := 20.0;  // 筛下流量 [立方米每小时] / the under sieve flow [cubic metre per hour]
    fQMin       : LREAL := 2.0;   // 流量下限（判据与除子域）[立方米每小时]，域 大于零 / the flow floor for the criteria and the divisor, domain above zero
    fWarnRatio  : LREAL := 1.5;   // 预警级比值阈 [无量纲]，域 大于 1 / the warning ratio threshold, above one
    fAlarmRatio : LREAL := 2.5;   // 报警级比值阈 [无量纲]，域 大于预警阈 / the alarm ratio threshold, above the warning one
    fCleanRatio : LREAL := 1.2;   // 清洁态比值上限（学习判据）[无量纲] / the clean ratio ceiling for learning
    tLearnWin   : TIME := T#60S;  // 清洁态学习持续窗 [毫秒]，域 大于零 / the clean learning dwell window [millisecond], domain above zero
END_VAR
VAR_OUTPUT
    fClogIdx    : LREAL := 1.0; // 堵塞指数（相对基准）[无量纲] / the clog index relative to the baseline
    fTrendSlope : LREAL := 0.0; // 8 点趋势斜率 [指数每拍] / the eight point trend slope [index per scan]
    ePhase      : E_DL_SscPhase := E_DL_SscPhase.eIdle; // 相位出口 [枚举] / phase outlet [enum]
    eFault      : E_DL_SscFault := E_DL_SscFault.eNone; // 成因出口，锁存回放 [枚举] / cause outlet replayed from the latch [enum]
    bError      : BOOL := FALSE; // 故障锁存标志 [-] / fault latch flag
END_VAR
VAR
    rtReset  : R_TRIG; // 复位沿检测，段 0 无条件刷新 / reset edge, refreshed unconditionally in segment zero
    rtLearn  : R_TRIG; // 学习窗到时沿检测，段 0 无条件刷新 / the learning window edge, refreshed unconditionally in segment zero
    tonLearn : TON;    // 清洁态学习持续窗（自清洁判据驱动，非错峰窗，无自复位需求）/ the clean learning dwell window
    _ePhase  : E_DL_SscPhase := E_DL_SscPhase.eIdle; // 内部相位，CASE 唯一写入目标 / internal phase, the only CASE write target
    _eFaulC  : E_DL_SscFault := E_DL_SscFault.eNone; // 故障级成因，锁存至复位沿 / fault cause, latched until the reset edge
    _bFault  : BOOL := FALSE; // 故障锁存位 [-] / fault latch bit
    _bInit   : BOOL := FALSE; // 首扫初始化完成标志（R310）/ first scan initialisation flag
    _bInOk   : BOOL := FALSE; // 两输入均有限 [-] / both inputs are finite
    _bCfgOk  : BOOL := FALSE; // 组态参数域内 [-] / the configuration is inside the domain
    _bBad    : BOOL := FALSE; // 传感器无效锁存 [-] / the sensor bad latch
    _bFlowLo : BOOL := FALSE; // 流量损失迟滞锁存 [-] / the flow loss hysteresis latch
    _bWarn   : BOOL := FALSE; // 预警迟滞锁存 [-] / the warning hysteresis latch
    _bAlarm  : BOOL := FALSE; // 报警迟滞锁存 [-] / the alarm hysteresis latch
    _bClean  : BOOL := FALSE; // 清洁态判定 [-] / the clean state verdict
    _nHead   : INT := 0;      // 环窗最近样本槽位（1 起）[槽号] / the newest ring slot, one based
    _nFill   : INT := 0;      // 环窗已填样本数 [个] / the ring fill count
    _nIdx    : INT := 1;      // 时间序遍历槽位 [槽号] / the time order traversal slot
    _nK      : INT := 0;      // 时间序遍历序号 [序号] / the time order ordinal
    _nGuard  : INT := 0;      // 遍历守护计数 [次] / the traversal guard [count]
    _fIdxRaw : LREAL := 0.0;  // 原始堵塞指数（dP / q²）[无量纲] / the raw clog index, dP over q squared
    _fSev    : LREAL := 0.0;  // 严重度（对基准比值）[无量纲] / the severity against the baseline
    _fSumX   : LREAL := 0.0;  // 最小二乘 Σx [无量纲] / the least squares sum of x
    _fSumY   : LREAL := 0.0;  // 最小二乘 Σy [无量纲] / the least squares sum of y
    _fSumXY  : LREAL := 0.0;  // 最小二乘 Σxy [无量纲] / the least squares sum of x times y
    _fNum    : LREAL := 0.0;  // 斜率分子 [无量纲] / the slope numerator
    _afIdx   : ARRAY[1..8] OF LREAL := [8(0.0)]; // 环窗堵塞指数缓存 [无量纲] / the ring of clog indices
END_VAR

// 段 0｜定时器与沿检测无条件周期刷新（禁入分支），IN 只串状态闸（FB50-1）/ segment 0, unconditional refresh with the state gates on IN only
rtReset(CLK := bReset); // 复位沿无条件刷新 / unconditional refresh of the reset edge
tonLearn(IN := _bClean AND (_ePhase = E_DL_SscPhase.eRun) AND (NOT _bFault) AND (NOT _bFlowLo) AND (NOT _bWarn) AND (NOT _bAlarm), PT := tLearnWin); // 清洁态学习窗 / the clean learning window
rtLearn(CLK := tonLearn.Q); // 学习窗到时沿 / the learning window edge

// 段 1｜首扫初始化（R310）/ segment 1, first scan initialisation
IF NOT _bInit THEN // 首扫一拍 / the very first scan
    _bInit := TRUE; // 置首扫完成标志 / raise the first scan flag
    _ePhase := E_DL_SscPhase.eRun; // 相位从运行起步 / the phase starts in run
    _eFaulC := E_DL_SscFault.eNone; // 故障级成因清零 / clear the fault cause
    _bFault := FALSE; // 故障锁存清零 / clear the fault latch
    _nHead := 0; // 环窗无样本 / the ring holds no sample
    _nFill := 0; // 环窗计数清零 / clear the ring count
END_IF

// 段 2｜复位沿作用域：清锁存 / 迁相位 / 清环窗与基准（三项逐项声明）/ segment 2, reset edge scope declared item by item
IF rtReset.Q THEN // 复位沿 / the reset edge
    _bFault := FALSE; // 作用域一：清故障锁存 / scope one, clear the fault latch
    _eFaulC := E_DL_SscFault.eNone; // 作用域一：清故障级成因 / scope one, clear the fault cause
    _bFlowLo := FALSE; // 作用域一：清流量损失迟滞 / scope one, clear the flow loss latch
    _bWarn := FALSE; // 作用域一：清预警迟滞 / scope one, clear the warning latch
    _bAlarm := FALSE; // 作用域一：清报警迟滞 / scope one, clear the alarm latch
    _bBad := FALSE; // 作用域一：清传感器锁存 / scope one, clear the sensor latch
    _ePhase := E_DL_SscPhase.eRun; // 作用域二：迁回运行相 / scope two, migrate back to run
    _nHead := 0; // 作用域三：清环窗槽位 / scope three, clear the ring slot
    _nFill := 0; // 作用域三：清环窗计数 / scope three, clear the ring count
    fClogIdx := 1.0; // 作用域三：指数回归基准水平 / scope three, the index returns to the baseline level
END_IF

// 段 3｜组态与输入域闸（R151 全覆盖）/ segment 3, the configuration and input domain gates
_bInOk := (fDp = fDp) AND ((fDp - fDp) = (fDp - fDp)) AND (fQ = fQ) AND ((fQ - fQ) = (fQ - fQ)); // 两输入有限性 / finiteness of both inputs
_bCfgOk := (fQMin > 0.0) AND (fQMin = fQMin) AND (fWarnRatio > 1.0) AND (fWarnRatio = fWarnRatio) AND (fAlarmRatio > fWarnRatio) AND (fAlarmRatio = fAlarmRatio) AND (fCleanRatio > 1.0) AND (fCleanRatio <= fWarnRatio) AND (fCleanRatio = fCleanRatio) AND (tLearnWin > T#0S); // 组态参数域判定 / the configuration domain verdict
IF (NOT _bInOk) OR (NOT _bCfgOk) THEN // 输入非有限或组态非法 / a non finite input or an illegal configuration
    IF NOT _bBad THEN // 未锁存才置 / set only while unlatched
        _bBad := TRUE; // 置传感器无效锁存 / raise the sensor bad latch
    END_IF
END_IF

// 段 4｜本拍指数计算与环窗写入 / segment 4, the per scan index computation and the ring write
_fIdxRaw := 0.0; // 原始指数预置零 / preset the raw index to zero
IF _bInOk AND (fQ > fQMin) THEN // 流量高于下限才可算（除子域闸）/ the index needs the flow above the floor
    _fIdxRaw := fDp / (fQ * fQ); // 原始堵塞指数，除子为流量平方已证超阈 / the raw index with the proven squared flow divisor
END_IF
IF (_nFill < 8) OR (_nHead < 8) THEN // 槽位推进（未满顺填，已满环回钳 1..8）/ advance the slot with the wrap clamp
    _nHead := _nHead + 1; // 槽位前移 / advance the slot
    IF _nHead > 8 THEN // 越过上界 / past the upper bound
        _nHead := 1; // 回钳到一号槽 / clamp back to slot one
    END_IF
    IF _nFill < 8 THEN // 未满顺填 / fill while not full
        _nFill := _nFill + 1; // 计数递增 / increment the count
    END_IF
    _afIdx[_nHead] := _fIdxRaw; // 指数入环窗 / store the index
END_IF

// 段 5｜时间序环窗遍历：最小二乘斜率（R194：自最旧样本起）/ segment 5, the time order traversal for the least squares slope
_fSumX := 0.0; // Σx 清零 / clear the sum of x
_fSumY := 0.0; // Σy 清零 / clear the sum of y
_fSumXY := 0.0; // Σxy 清零 / clear the sum of xy
fTrendSlope := 0.0; // 斜率输出每拍预置零（样本不足时保持零，最小二乘仅在窗内覆盖）/ preset the slope outlet to zero, recomputed only when enough samples
IF _nFill >= 2 THEN // 至少两点才可算斜率 / the slope needs at least two points
    _nK := 1; // 时间序序号起步（1 = 最旧样本）/ start the time order ordinal at the oldest
    _nGuard := 0; // 守护清零 / clear the guard
    WHILE (_nK <= _nFill) AND (_nGuard < 16) DO // 时间序遍历，守护为两倍容量 / the time order traversal with a twice capacity guard
        _nGuard := _nGuard + 1; // 守护递增 / increment the guard
        _nIdx := _nHead - _nFill + _nK; // 时间序槽位 / the slot in time order
        IF _nIdx < 1 THEN // 越过下界 / below the lower bound
            _nIdx := _nIdx + 8; // 单次回绕补齐 / a single wrap restores the order
        END_IF
        _fSumX := _fSumX + INT_TO_LREAL(_nK - 1); // x = 0..7 / the x ordinal from zero
        _fSumY := _fSumY + _afIdx[_nIdx]; // y 累计 / accumulate y
        _fSumXY := _fSumXY + INT_TO_LREAL(_nK - 1) * _afIdx[_nIdx]; // xy 累计 / accumulate xy
        _nK := _nK + 1; // 序号递增 / increment the ordinal
    END_WHILE
    _fNum := 8.0 * _fSumXY - _fSumX * _fSumY; // 斜率分子 / the slope numerator
    fTrendSlope := _fNum / 336.0; // 最小二乘斜率，分母 8·140 - 28² = 336 结构性非零（R63 反算留档）/ the slope, the denominator is structurally non zero
END_IF

// 段 6｜严重度计算（对时间序最旧样本 = 学习基准）/ segment 6, the severity against the oldest sample as the learned baseline
IF _nFill >= 1 THEN // 有样本 / a sample exists
    _nIdx := _nHead - _nFill + 1; // 时间序最旧槽位（学习基准）/ the oldest slot, the learned baseline
    IF _nIdx < 1 THEN // 越过下界 / below the lower bound
        _nIdx := _nIdx + 8; // 单次回绕 / a single wrap
    END_IF
    IF _afIdx[_nIdx] > 1.0E-9 THEN // 基准指数可用（除子域闸）/ the baseline is usable
        fClogIdx := _afIdx[_nHead] / _afIdx[_nIdx]; // 堵塞指数 = 当前 / 学习基准 / the clog index, the current over the learned baseline
        _fSev := fClogIdx; // 严重度同源 / the severity shares the source
    ELSE // 基准指数近零 / the baseline is near zero
        fClogIdx := 1.0; // 指数回归基准 / the index returns to the baseline
        _fSev := 1.0; // 严重度记一 / the severity is one
    END_IF
ELSE // 无样本 / no sample
    fClogIdx := 1.0; // 指数回归基准 / the index returns to the baseline
    _fSev := 1.0; // 严重度记一 / the severity is one
END_IF
_bClean := (_fSev <= fCleanRatio) AND (fQ > fQMin) AND _bInOk; // 清洁态判定 / the clean state verdict
IF _fSev > fAlarmRatio THEN // 报警级进入判据 / the alarm entry criterion
    _bAlarm := TRUE; // 置报警迟滞 / raise the alarm latch
    _bWarn := TRUE; // 报警级蕴含预警级 / the alarm implies the warning
ELSIF _fSev < fWarnRatio - 0.1 THEN // 报警级退出判据（迟滞收窄）/ the alarm exit criterion with the narrowed band
    _bAlarm := FALSE; // 清报警迟滞 / clear the alarm latch
END_IF
IF (_fSev > fWarnRatio) AND (NOT _bAlarm) THEN // 预警级进入判据 / the warning entry criterion
    _bWarn := TRUE; // 置预警迟滞 / raise the warning latch
ELSIF _fSev < fWarnRatio - 0.1 THEN // 预警级退出判据（迟滞收窄）/ the warning exit criterion
    _bWarn := FALSE; // 清预警迟滞 / clear the warning latch
END_IF
IF fQ <= fQMin THEN // 流量损失进入判据 / the flow loss entry criterion
    _bFlowLo := TRUE; // 置流量损失迟滞 / raise the flow loss latch
ELSIF fQ > fQMin * 1.2 THEN // 流量损失退出判据（迟滞收窄）/ the flow loss exit criterion
    _bFlowLo := FALSE; // 清流量损失迟滞 / clear the flow loss latch
END_IF

// 段 7｜相位机：ENUM + CASE，含 ELSE 非法相位兜底（R128）/ segment 7, the phase machine with an ELSE fallback
CASE _ePhase OF
E_DL_SscPhase.eIdle: // 未使能相 / the disabled phase
    IF bEnable AND (NOT _bFault) THEN // 使能且无故障 / enabled and unfaulted
        _ePhase := E_DL_SscPhase.eRun; // 迁运行相 / migrate to run
    END_IF

E_DL_SscPhase.eRun: // 运行相：判级分派（优先级：传感器 > 流量损失 > 报警 > 预警）与学习更新 / the run phase, the dispatch and the learning
    IF NOT bEnable THEN // 失能 / disabled
        _ePhase := E_DL_SscPhase.eIdle; // 迁未使能相 / migrate to idle
    ELSIF _bBad OR _bFlowLo OR _bAlarm OR _bWarn THEN // 存在活跃迟滞锁存 / an active latch exists
        _bFault := TRUE; // 置故障锁存 / raise the fault latch
        IF _bBad THEN // 传感器非有限优先 / the sensor takes the top priority
            _eFaulC := E_DL_SscFault.eSensorBad; // 故障级成因（R45 配对 bError）/ the fault cause paired with bError
        ELSIF _bFlowLo THEN // 流量损失次优先 / the flow loss follows
            _eFaulC := E_DL_SscFault.eFlowLoss; // 故障级成因（R45 配对 bError）/ the fault cause paired with bError
        ELSIF _bAlarm THEN // 报警级再次优先（R190 独立成因）/ the alarm grade, an independent cause
            _eFaulC := E_DL_SscFault.eClogAlarm; // 故障级成因（R45 配对 bError）/ the fault cause paired with bError
        ELSE // 预警级（R190 独立成因）/ the warning grade, an independent cause
            _eFaulC := E_DL_SscFault.eClogWarn; // 故障级成因（R45 配对 bError）/ the fault cause paired with bError
        END_IF
        _ePhase := E_DL_SscPhase.eFault; // 迁故障相 / migrate to the fault phase
    ELSE // 正常运行 / the normal running
        _eFaulC := E_DL_SscFault.eNone; // 成因清零 / clear the cause
    END_IF

E_DL_SscPhase.eFault: // 故障相：锁存回放，迟滞自愈解除后回运行 / the fault phase, the latches self heal and return to run
    IF bEnable AND (NOT _bBad) AND (NOT _bFlowLo) AND (NOT _bAlarm) AND (NOT _bWarn) THEN // 全部迟滞已解除 / every latch has cleared
        _bFault := FALSE; // 清故障锁存（自愈路径，R152）/ clear the fault latch, the self healing path
        _eFaulC := E_DL_SscFault.eNone; // 成因清零 / clear the cause
        _ePhase := E_DL_SscPhase.eRun; // 迁回运行相 / migrate back to run
    ELSIF NOT bEnable THEN // 失能 / disabled
        _ePhase := E_DL_SscPhase.eIdle; // 迁未使能相 / migrate to idle
    END_IF

ELSE // 非法相位兜底（R128）/ the illegal phase fallback
    _bFault := TRUE; // 置故障锁存 / raise the fault latch
    _eFaulC := E_DL_SscFault.ePhaseBad; // 故障级成因（R45 配对 bError）/ the fault cause paired with bError
    _ePhase := E_DL_SscPhase.eFault; // 迁故障相 / migrate to the fault phase
END_CASE

// 段 8｜学习更新与统一出口 / segment 8, the learning update and the unified outlet
IF rtLearn.Q THEN // 学习窗到时沿 / the learning edge
    _nIdx := _nHead - _nFill + 1; // 时间序最旧槽位 / the oldest slot in time order
    IF _nIdx < 1 THEN // 越过下界 / below the lower bound
        _nIdx := _nIdx + 8; // 单次回绕 / a single wrap
    END_IF
    _afIdx[_nIdx] := _afIdx[_nHead]; // 基准更新：最旧样本改写为当前指数 / the baseline update, the oldest slot takes the current index
END_IF
IF _bFault THEN // 故障锁存优先 / the fault latch takes priority
    eFault := _eFaulC; // 故障级成因锁存回放（R152）/ the fault cause replayed from the latch
ELSE
    eFault := E_DL_SscFault.eNone; // 无锁存即无成因 / no latch, no cause
END_IF
ePhase := _ePhase; // 相位出口单点映射 / single point phase outlet mapping
bError := _bFault; // 故障标志与锁存位同源 / the fault flag shares the latch source
END_FUNCTION_BLOCK

(* ---- FB_DL_SpliceCountdownCtrl.st ---- *)
(*
  DL Factory R83 | FB_DL_SpliceCountdownCtrl
  功能：按当前卷径反算接卷剩余米数，用两段阈值加回差带输出预警与报警。
  开源溯源：无（clean-room 自研，依据公开工艺公式，来源=行业通用公式，许可证=MIT，借鉴点=公式结构）
  规则：R1-R21 全遵守
*)
FUNCTION_BLOCK FB_DL_SpliceCountdownCtrl
VAR_INPUT
    fRollDiaMm  : REAL; // 当前卷径 [mm] / Current roll diameter [mm]
    fCoreDiaMm  : REAL; // 卷芯直径 [mm] / Core diameter [mm]
    fWebThickMm : REAL; // 料带厚度 [mm] / Web thickness [mm]
    fWarnM      : REAL; // 预警剩余米数阈值 [m] / Warning remaining threshold [m]
    fAlarmM     : REAL; // 报警剩余米数阈值 [m] / Alarm remaining threshold [m]
    bReset      : BOOL; // 复位：清故障码 / Reset: clear error code
END_VAR
VAR_OUTPUT
    fRemainM : REAL; // 剩余料长 [m] / Remaining web length [m]
    xWarn    : BOOL; // 预警输出（可准备换卷）/ Warning output (prepare splice)
    xAlarm   : BOOL; // 报警输出（立即接卷）/ Alarm output (splice now)
    iErrCode : INT;  // 错误码，0=无错 / Error code, 0 = no error
END_VAR
VAR
    fR2Mm : REAL; // 半径平方差（R²-r²）[mm²] / Radius-square difference [mm^2]
END_VAR

// ---------- 出口预置：信息位每拍重算（R187/R256） ----------
fRemainM := 0.0;                      // 剩余料长预置零 [m] / Remaining length preset zero
xWarn    := FALSE; xAlarm := FALSE;   // 双标志预置 FALSE（名实双出口同源，R191）
IF bReset THEN iErrCode := 0; END_IF  // 故障码唯一清除边：bReset 上升沿（R188）

// ---------- 非有限 + 量纲次序 + 分母零闸：一次拦截（R4/R20/R21） ----------
IF NOT (fRollDiaMm > -1.0E30 AND fRollDiaMm < 1.0E30) OR NOT (fCoreDiaMm > -1.0E30 AND fCoreDiaMm < 1.0E30) OR NOT (fWebThickMm > -1.0E30 AND fWebThickMm < 1.0E30) OR NOT (fWarnM > -1.0E30 AND fWarnM < 1.0E30) OR NOT (fAlarmM > -1.0E30 AND fAlarmM < 1.0E30) OR fRollDiaMm <= fCoreDiaMm OR fWarnM <= fAlarmM OR ABS(fWebThickMm) <= 1.0E-9 THEN
    iErrCode := 9001;                 // 非有限/量纲越界/厚度零值统一码 / Non-finite, dimension, zero thickness
    RETURN;                           // 故障拍不出报警，交由上层按码处置 / Fault cycle emits no alarm
END_IF

// ---------- 剩余料长：L = π × (R² - r²) / t，mm ÷ 1000 换算为 m ----------
fR2Mm    := (fRollDiaMm * fRollDiaMm - fCoreDiaMm * fCoreDiaMm) / 4.0; // 半径平方差 [mm²]
fRemainM := 3.14159265358979 * fR2Mm / fWebThickMm / 1000.0;           // 剩余料长 [m]

// ---------- 两段阈值 + 0.5 m 回差带：进入即置，退出须越过阈值加回差 ----------
IF fRemainM <= fWarnM THEN xWarn := TRUE; END_IF                          // 进入预警带 / Enter warning band
IF fRemainM <= fAlarmM THEN xAlarm := TRUE; xWarn := TRUE; END_IF         // 报警带蕴含预警（R191 名实双置）
IF fRemainM > fWarnM + 0.5 THEN xWarn := FALSE; xAlarm := FALSE; END_IF   // 越过回差带回退 / Release past hysteresis
END_FUNCTION_BLOCK
